// ---- VISUs/Carrousel.TcVIS
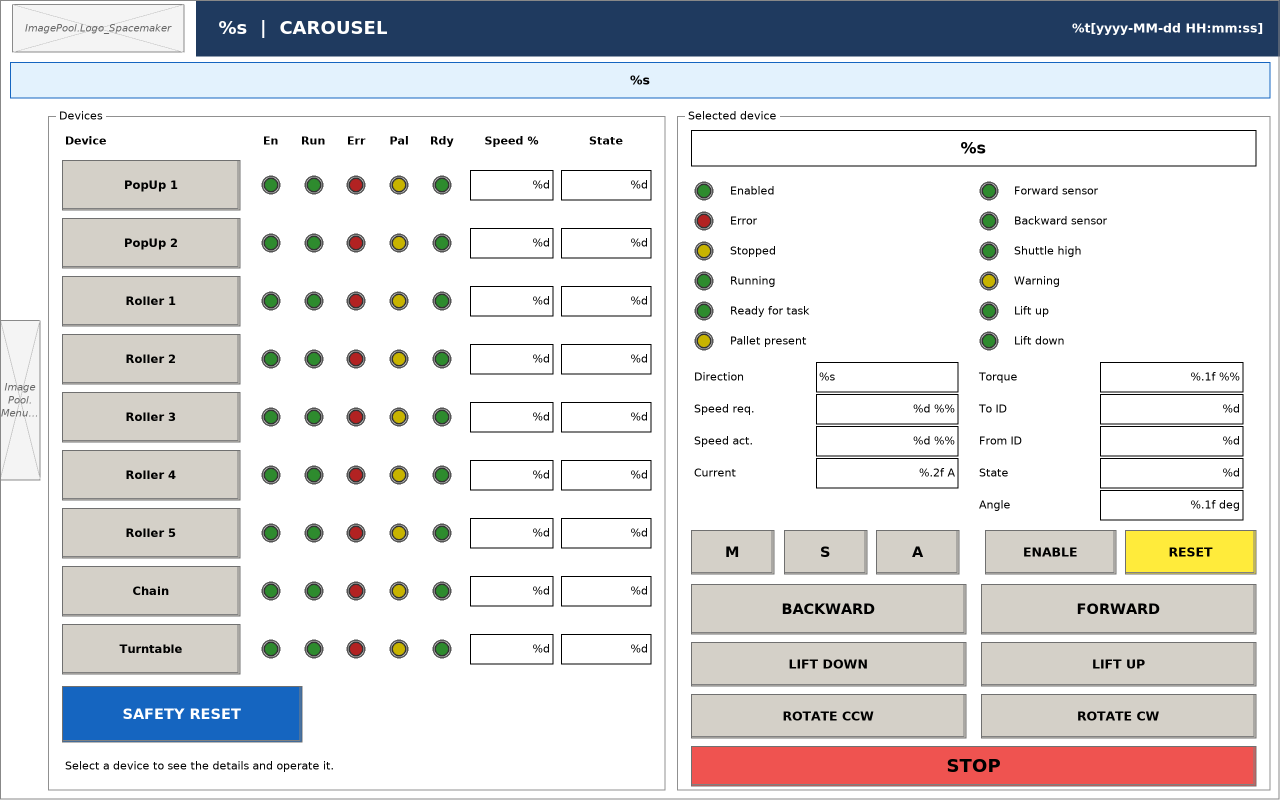
VISUALIZATION Carrousel  // 1280x800
    Rectangle (0,0 196x56)
        OnMouseClick: change screen: Main
    Image (12,4 172x48), image: ImagePool.Logo_Spacemaker
        OnMouseClick: change screen: Main
    Rectangle (196,0 1084x56), "%s | CAROUSEL", text variable: GVL_HMI_System.stStatus.sSystemName
    Rectangle (930,8 336x40), "%t[yyyy-MM-dd HH:mm:ss]", text variable: GVL_HMI_System.stStatus.dtNow
    Rectangle (10,62 1260x36), "%s", text variable: GVL_HMI_System.stStatus.sMessage, colour toggle: GVL_HMI_System.stStatus.bMessageAlarm
    GroupBox (48,108 617x682), "Devices"
    Rectangle (62,128 178x26), "Device"
    Rectangle (250,128 42x26), "En"
    Rectangle (292,128 43x26), "Run"
    Rectangle (335,128 43x26), "Err"
    Rectangle (378,128 43x26), "Pal"
    Rectangle (421,128 42x26), "Rdy"
    Rectangle (470,128 83x26), "Speed %"
    Rectangle (561,128 90x26), "State"
    Button (62,160 178x50), "PopUp 1", colour toggle: GVL_HMI_Carousel.astDevice[1].bSelected
        OnMouseClick: execute { GVL_HMI_Carousel.uiSelected := 1; }
    Lamp1 (260,174 22x22), variable: GVL_HMI_Carousel.astDevice[1].bEnabled, style: Lamp-Lamp1-Green
    Lamp1 (303,174 22x22), variable: GVL_HMI_Carousel.astDevice[1].bRunning, style: Lamp-Lamp1-Green
    Lamp1 (345,174 22x22), variable: GVL_HMI_Carousel.astDevice[1].bError, style: Lamp-Lamp1-Red
    Lamp1 (388,174 22x22), variable: GVL_HMI_Carousel.astDevice[1].bOccupied, style: Lamp-Lamp1-Yellow
    Lamp1 (431,174 22x22), variable: GVL_HMI_Carousel.astDevice[1].bReadyForTask, style: Lamp-Lamp1-Green
    Rectangle (470,170 83x30), "%d", text variable: GVL_HMI_Carousel.astDevice[1].iSpeedActual_pct
    Rectangle (561,170 90x30), "%d", text variable: GVL_HMI_Carousel.astDevice[1].uiStateMachine
    Button (62,218 178x50), "PopUp 2", colour toggle: GVL_HMI_Carousel.astDevice[2].bSelected
        OnMouseClick: execute { GVL_HMI_Carousel.uiSelected := 2; }
    Lamp1 (260,232 22x22), variable: GVL_HMI_Carousel.astDevice[2].bEnabled, style: Lamp-Lamp1-Green
    Lamp1 (303,232 22x22), variable: GVL_HMI_Carousel.astDevice[2].bRunning, style: Lamp-Lamp1-Green
    Lamp1 (345,232 22x22), variable: GVL_HMI_Carousel.astDevice[2].bError, style: Lamp-Lamp1-Red
    Lamp1 (388,232 22x22), variable: GVL_HMI_Carousel.astDevice[2].bOccupied, style: Lamp-Lamp1-Yellow
    Lamp1 (431,232 22x22), variable: GVL_HMI_Carousel.astDevice[2].bReadyForTask, style: Lamp-Lamp1-Green
    Rectangle (470,228 83x30), "%d", text variable: GVL_HMI_Carousel.astDevice[2].iSpeedActual_pct
    Rectangle (561,228 90x30), "%d", text variable: GVL_HMI_Carousel.astDevice[2].uiStateMachine
    Button (62,276 178x50), "Roller 1", colour toggle: GVL_HMI_Carousel.astDevice[3].bSelected
        OnMouseClick: execute { GVL_HMI_Carousel.uiSelected := 3; }
    Lamp1 (260,290 22x22), variable: GVL_HMI_Carousel.astDevice[3].bEnabled, style: Lamp-Lamp1-Green
    Lamp1 (303,290 22x22), variable: GVL_HMI_Carousel.astDevice[3].bRunning, style: Lamp-Lamp1-Green
    Lamp1 (345,290 22x22), variable: GVL_HMI_Carousel.astDevice[3].bError, style: Lamp-Lamp1-Red
    Lamp1 (388,290 22x22), variable: GVL_HMI_Carousel.astDevice[3].bOccupied, style: Lamp-Lamp1-Yellow
    Lamp1 (431,290 22x22), variable: GVL_HMI_Carousel.astDevice[3].bReadyForTask, style: Lamp-Lamp1-Green
    Rectangle (470,286 83x30), "%d", text variable: GVL_HMI_Carousel.astDevice[3].iSpeedActual_pct
    Rectangle (561,286 90x30), "%d", text variable: GVL_HMI_Carousel.astDevice[3].uiStateMachine
    Button (62,334 178x50), "Roller 2", colour toggle: GVL_HMI_Carousel.astDevice[4].bSelected
        OnMouseClick: execute { GVL_HMI_Carousel.uiSelected := 4; }
    Lamp1 (260,348 22x22), variable: GVL_HMI_Carousel.astDevice[4].bEnabled, style: Lamp-Lamp1-Green
    Lamp1 (303,348 22x22), variable: GVL_HMI_Carousel.astDevice[4].bRunning, style: Lamp-Lamp1-Green
    Lamp1 (345,348 22x22), variable: GVL_HMI_Carousel.astDevice[4].bError, style: Lamp-Lamp1-Red
    Lamp1 (388,348 22x22), variable: GVL_HMI_Carousel.astDevice[4].bOccupied, style: Lamp-Lamp1-Yellow
    Lamp1 (431,348 22x22), variable: GVL_HMI_Carousel.astDevice[4].bReadyForTask, style: Lamp-Lamp1-Green
    Rectangle (470,344 83x30), "%d", text variable: GVL_HMI_Carousel.astDevice[4].iSpeedActual_pct
    Rectangle (561,344 90x30), "%d", text variable: GVL_HMI_Carousel.astDevice[4].uiStateMachine
    Button (62,392 178x50), "Roller 3", colour toggle: GVL_HMI_Carousel.astDevice[5].bSelected
        OnMouseClick: execute { GVL_HMI_Carousel.uiSelected := 5; }
    Lamp1 (260,406 22x22), variable: GVL_HMI_Carousel.astDevice[5].bEnabled, style: Lamp-Lamp1-Green
    Lamp1 (303,406 22x22), variable: GVL_HMI_Carousel.astDevice[5].bRunning, style: Lamp-Lamp1-Green
    Lamp1 (345,406 22x22), variable: GVL_HMI_Carousel.astDevice[5].bError, style: Lamp-Lamp1-Red
    Lamp1 (388,406 22x22), variable: GVL_HMI_Carousel.astDevice[5].bOccupied, style: Lamp-Lamp1-Yellow
    Lamp1 (431,406 22x22), variable: GVL_HMI_Carousel.astDevice[5].bReadyForTask, style: Lamp-Lamp1-Green
    Rectangle (470,402 83x30), "%d", text variable: GVL_HMI_Carousel.astDevice[5].iSpeedActual_pct
    Rectangle (561,402 90x30), "%d", text variable: GVL_HMI_Carousel.astDevice[5].uiStateMachine
    Button (62,450 178x50), "Roller 4", colour toggle: GVL_HMI_Carousel.astDevice[6].bSelected
        OnMouseClick: execute { GVL_HMI_Carousel.uiSelected := 6; }
    Lamp1 (260,464 22x22), variable: GVL_HMI_Carousel.astDevice[6].bEnabled, style: Lamp-Lamp1-Green
    Lamp1 (303,464 22x22), variable: GVL_HMI_Carousel.astDevice[6].bRunning, style: Lamp-Lamp1-Green
    Lamp1 (345,464 22x22), variable: GVL_HMI_Carousel.astDevice[6].bError, style: Lamp-Lamp1-Red
    Lamp1 (388,464 22x22), variable: GVL_HMI_Carousel.astDevice[6].bOccupied, style: Lamp-Lamp1-Yellow
    Lamp1 (431,464 22x22), variable: GVL_HMI_Carousel.astDevice[6].bReadyForTask, style: Lamp-Lamp1-Green
    Rectangle (470,460 83x30), "%d", text variable: GVL_HMI_Carousel.astDevice[6].iSpeedActual_pct
    Rectangle (561,460 90x30), "%d", text variable: GVL_HMI_Carousel.astDevice[6].uiStateMachine
    Button (62,508 178x50), "Roller 5", colour toggle: GVL_HMI_Carousel.astDevice[7].bSelected
        OnMouseClick: execute { GVL_HMI_Carousel.uiSelected := 7; }
    Lamp1 (260,522 22x22), variable: GVL_HMI_Carousel.astDevice[7].bEnabled, style: Lamp-Lamp1-Green
    Lamp1 (303,522 22x22), variable: GVL_HMI_Carousel.astDevice[7].bRunning, style: Lamp-Lamp1-Green
    Lamp1 (345,522 22x22), variable: GVL_HMI_Carousel.astDevice[7].bError, style: Lamp-Lamp1-Red
    Lamp1 (388,522 22x22), variable: GVL_HMI_Carousel.astDevice[7].bOccupied, style: Lamp-Lamp1-Yellow
    Lamp1 (431,522 22x22), variable: GVL_HMI_Carousel.astDevice[7].bReadyForTask, style: Lamp-Lamp1-Green
    Rectangle (470,518 83x30), "%d", text variable: GVL_HMI_Carousel.astDevice[7].iSpeedActual_pct
    Rectangle (561,518 90x30), "%d", text variable: GVL_HMI_Carousel.astDevice[7].uiStateMachine
    Button (62,566 178x50), "Chain", colour toggle: GVL_HMI_Carousel.astDevice[8].bSelected
        OnMouseClick: execute { GVL_HMI_Carousel.uiSelected := 8; }
    Lamp1 (260,580 22x22), variable: GVL_HMI_Carousel.astDevice[8].bEnabled, style: Lamp-Lamp1-Green
    Lamp1 (303,580 22x22), variable: GVL_HMI_Carousel.astDevice[8].bRunning, style: Lamp-Lamp1-Green
    Lamp1 (345,580 22x22), variable: GVL_HMI_Carousel.astDevice[8].bError, style: Lamp-Lamp1-Red
    Lamp1 (388,580 22x22), variable: GVL_HMI_Carousel.astDevice[8].bOccupied, style: Lamp-Lamp1-Yellow
    Lamp1 (431,580 22x22), variable: GVL_HMI_Carousel.astDevice[8].bReadyForTask, style: Lamp-Lamp1-Green
    Rectangle (470,576 83x30), "%d", text variable: GVL_HMI_Carousel.astDevice[8].iSpeedActual_pct
    Rectangle (561,576 90x30), "%d", text variable: GVL_HMI_Carousel.astDevice[8].uiStateMachine
    Button (62,624 178x50), "Turntable", colour toggle: GVL_HMI_Carousel.astDevice[9].bSelected
        OnMouseClick: execute { GVL_HMI_Carousel.uiSelected := 9; }
    Lamp1 (260,638 22x22), variable: GVL_HMI_Carousel.astDevice[9].bEnabled, style: Lamp-Lamp1-Green
    Lamp1 (303,638 22x22), variable: GVL_HMI_Carousel.astDevice[9].bRunning, style: Lamp-Lamp1-Green
    Lamp1 (345,638 22x22), variable: GVL_HMI_Carousel.astDevice[9].bError, style: Lamp-Lamp1-Red
    Lamp1 (388,638 22x22), variable: GVL_HMI_Carousel.astDevice[9].bOccupied, style: Lamp-Lamp1-Yellow
    Lamp1 (431,638 22x22), variable: GVL_HMI_Carousel.astDevice[9].bReadyForTask, style: Lamp-Lamp1-Green
    Rectangle (470,634 83x30), "%d", text variable: GVL_HMI_Carousel.astDevice[9].iSpeedActual_pct
    Rectangle (561,634 90x30), "%d", text variable: GVL_HMI_Carousel.astDevice[9].uiStateMachine
    Rectangle (62,752 593x28), "Select a device to see the details and operate it."
    GroupBox (677,108 593x682), "Selected device"
    Rectangle (691,130 565x36), "%s", text variable: GVL_HMI_Carousel.stSelected.sName
    Lamp1 (693,180 22x22), variable: GVL_HMI_Carousel.stSelected.bEnabled, style: Lamp-Lamp1-Green
    Rectangle (727,176 201x30), "Enabled"
    Lamp1 (693,210 22x22), variable: GVL_HMI_Carousel.stSelected.bError, style: Lamp-Lamp1-Red
    Rectangle (727,206 201x30), "Error"
    Lamp1 (693,240 22x22), variable: GVL_HMI_Carousel.stSelected.bStopped, style: Lamp-Lamp1-Yellow
    Rectangle (727,236 201x30), "Stopped"
    Lamp1 (693,270 22x22), variable: GVL_HMI_Carousel.stSelected.bRunning, style: Lamp-Lamp1-Green
    Rectangle (727,266 201x30), "Running"
    Lamp1 (693,300 22x22), variable: GVL_HMI_Carousel.stSelected.bReadyForTask, style: Lamp-Lamp1-Green
    Rectangle (727,296 201x30), "Ready for task"
    Lamp1 (693,330 22x22), variable: GVL_HMI_Carousel.stSelected.bOccupied, style: Lamp-Lamp1-Yellow
    Rectangle (727,326 201x30), "Pallet present"
    Lamp1 (978,180 22x22), variable: GVL_HMI_Carousel.stSelected.bForwardSensor, style: Lamp-Lamp1-Green
    Rectangle (1011,176 202x30), "Forward sensor"
    Lamp1 (978,210 22x22), variable: GVL_HMI_Carousel.stSelected.bBackwardSensor, style: Lamp-Lamp1-Green
    Rectangle (1011,206 202x30), "Backward sensor"
    Lamp1 (978,240 22x22), variable: GVL_HMI_Carousel.stSelected.bShuttleHigh, style: Lamp-Lamp1-Green
    Rectangle (1011,236 202x30), "Shuttle high"
    Lamp1 (978,270 22x22), variable: GVL_HMI_Carousel.stSelected.bWarning, style: Lamp-Lamp1-Yellow
    Rectangle (1011,266 202x30), "Warning"
    Lamp1 (978,300 22x22), variable: GVL_HMI_Carousel.stSelected.bLiftUp, style: Lamp-Lamp1-Green
    Rectangle (1011,296 202x30), "Lift up"
    Lamp1 (978,330 22x22), variable: GVL_HMI_Carousel.stSelected.bLiftDown, style: Lamp-Lamp1-Green
    Rectangle (1011,326 202x30), "Lift down"
    Rectangle (691,362 119x30), "Direction"
    Rectangle (816,362 142x30), "%s", text variable: GVL_HMI_Carousel.stSelected.sMotorDirection
    Rectangle (691,394 119x30), "Speed req."
    Rectangle (816,394 142x30), "%d %%", text variable: GVL_HMI_Carousel.stSelected.iSpeedRequested_pct
    Rectangle (691,426 119x30), "Speed act."
    Rectangle (816,426 142x30), "%d %%", text variable: GVL_HMI_Carousel.stSelected.iSpeedActual_pct
    Rectangle (691,458 119x30), "Current"
    Rectangle (816,458 142x30), "%.2f A", text variable: GVL_HMI_Carousel.stSelected.rCurrent_A
    Rectangle (976,362 118x30), "Torque"
    Rectangle (1100,362 143x30), "%.1f %%", text variable: GVL_HMI_Carousel.stSelected.rTorque_pct
    Rectangle (976,394 118x30), "To ID"
    Rectangle (1100,394 143x30), "%d", text variable: GVL_HMI_Carousel.stSelected.diTransferToId
    Rectangle (976,426 118x30), "From ID"
    Rectangle (1100,426 143x30), "%d", text variable: GVL_HMI_Carousel.stSelected.diTransferFromId
    Rectangle (976,458 118x30), "State"
    Rectangle (1100,458 143x30), "%d", text variable: GVL_HMI_Carousel.stSelected.uiStateMachine
    Rectangle (976,490 118x30), "Angle"
    Rectangle (1100,490 143x30), "%.1f deg", text variable: GVL_HMI_Carousel.stSelected.rAngle_deg
    Button (691,530 83x44), "M", colour toggle: GVL_HMI_Carousel.stSelected.bModeManual
        tap GVL_HMI_Carousel.stCommand.bModeManual p3779583253=TRUE
    Button (784,530 83x44), "S", colour toggle: GVL_HMI_Carousel.stSelected.bModeSemi
        tap GVL_HMI_Carousel.stCommand.bModeSemi p3779583253=TRUE
    Button (876,530 83x44), "A", colour toggle: GVL_HMI_Carousel.stSelected.bModeAuto
        tap GVL_HMI_Carousel.stCommand.bModeAuto p3779583253=TRUE
    Button (985,530 131x44), "ENABLE", colour toggle: GVL_HMI_Carousel.stSelected.bEnabled
        tap GVL_HMI_Carousel.stCommand.bEnable p3779583253=TRUE
    Button (1125,530 131x44), "RESET"
        tap GVL_HMI_Carousel.stCommand.bReset p3779583253=TRUE
    Button (691,584 275x50), "BACKWARD", input disabled if: NOT GVL_HMI_Carousel.stSelected.bModeManual
        tap GVL_HMI_Carousel.stCommand.bJogBackward p3779583253=TRUE
    Button (981,584 275x50), "FORWARD", input disabled if: NOT GVL_HMI_Carousel.stSelected.bModeManual
        tap GVL_HMI_Carousel.stCommand.bJogForward p3779583253=TRUE
    Button (691,642 275x44), "LIFT DOWN", input disabled if: NOT GVL_HMI_Carousel.stSelected.bHasLift
        tap GVL_HMI_Carousel.stCommand.bLiftDown p3779583253=TRUE
    Button (981,642 275x44), "LIFT UP", input disabled if: NOT GVL_HMI_Carousel.stSelected.bHasLift
        tap GVL_HMI_Carousel.stCommand.bLiftUp p3779583253=TRUE
    Button (691,694 275x44), "ROTATE CCW", input disabled if: NOT GVL_HMI_Carousel.stSelected.bHasRotation
        tap GVL_HMI_Carousel.stCommand.bRotateCcw p3779583253=TRUE
    Button (981,694 275x44), "ROTATE CW", input disabled if: NOT GVL_HMI_Carousel.stSelected.bHasRotation
        tap GVL_HMI_Carousel.stCommand.bRotateCw p3779583253=TRUE
    Button (691,746 565x40), "STOP"
        tap GVL_HMI_Carousel.stCommand.bStop p3779583253=TRUE
    Rectangle (0,320 40x160)
        OnMouseClick: OpenDialog Dialog=Dialog, OpenModal=True, PositionX=0, PositionY=0
        OnMouseEnter: OpenDialog Dialog=Dialog, OpenModal=True, PositionX=0, PositionY=0
    Image (0,320 40x160), image: ImagePool.Menu_Tab
        OnMouseClick: OpenDialog Dialog=Dialog, OpenModal=True, PositionX=0, PositionY=0
        OnMouseEnter: OpenDialog Dialog=Dialog, OpenModal=True, PositionX=0, PositionY=0
    Button (62,686 240x56), "SAFETY RESET", colour toggle: GVL_HMI_System.stStatus.bSafetyResetActive
        tap GVL_HMI_System.stCommand.bSafetyReset p3779583253=TRUE
END_VISUALIZATION

// ---- VISUs/CNV.TcVIS
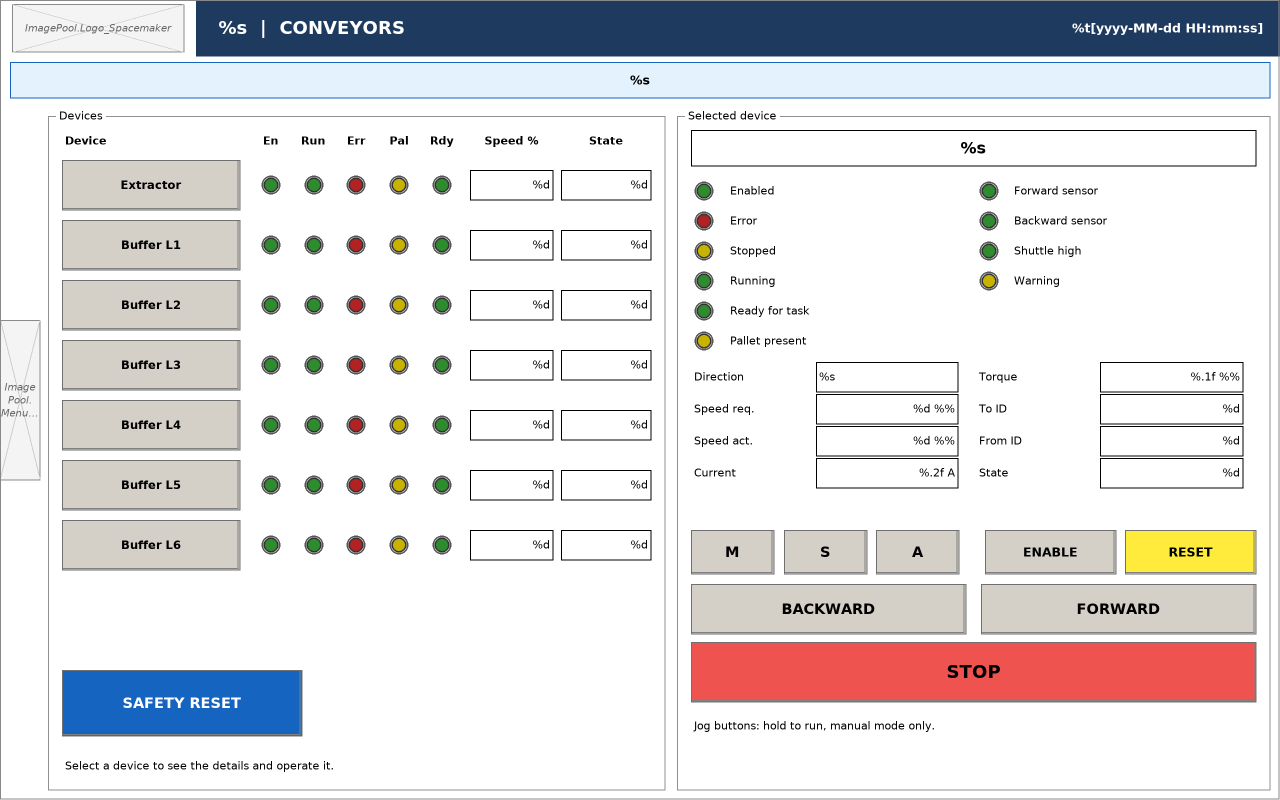
VISUALIZATION CNV  // 1280x800
    Rectangle (0,0 196x56)
        OnMouseClick: change screen: Main
    Image (12,4 172x48), image: ImagePool.Logo_Spacemaker
        OnMouseClick: change screen: Main
    Rectangle (196,0 1084x56), "%s | CONVEYORS", text variable: GVL_HMI_System.stStatus.sSystemName
    Rectangle (930,8 336x40), "%t[yyyy-MM-dd HH:mm:ss]", text variable: GVL_HMI_System.stStatus.dtNow
    Rectangle (10,62 1260x36), "%s", text variable: GVL_HMI_System.stStatus.sMessage, colour toggle: GVL_HMI_System.stStatus.bMessageAlarm
    GroupBox (48,108 617x682), "Devices"
    Rectangle (62,128 178x26), "Device"
    Rectangle (250,128 42x26), "En"
    Rectangle (292,128 43x26), "Run"
    Rectangle (335,128 43x26), "Err"
    Rectangle (378,128 43x26), "Pal"
    Rectangle (421,128 42x26), "Rdy"
    Rectangle (470,128 83x26), "Speed %"
    Rectangle (561,128 90x26), "State"
    Button (62,160 178x50), "Extractor", colour toggle: GVL_HMI_CNV.astConveyor[0].bSelected
        OnMouseClick: execute { GVL_HMI_CNV.uiSelected := 0; }
    Lamp1 (260,174 22x22), variable: GVL_HMI_CNV.astConveyor[0].bEnabled, style: Lamp-Lamp1-Green
    Lamp1 (303,174 22x22), variable: GVL_HMI_CNV.astConveyor[0].bRunning, style: Lamp-Lamp1-Green
    Lamp1 (345,174 22x22), variable: GVL_HMI_CNV.astConveyor[0].bError, style: Lamp-Lamp1-Red
    Lamp1 (388,174 22x22), variable: GVL_HMI_CNV.astConveyor[0].bOccupied, style: Lamp-Lamp1-Yellow
    Lamp1 (431,174 22x22), variable: GVL_HMI_CNV.astConveyor[0].bReadyForTask, style: Lamp-Lamp1-Green
    Rectangle (470,170 83x30), "%d", text variable: GVL_HMI_CNV.astConveyor[0].iSpeedActual_pct
    Rectangle (561,170 90x30), "%d", text variable: GVL_HMI_CNV.astConveyor[0].uiStateMachine
    Button (62,220 178x50), "Buffer L1", colour toggle: GVL_HMI_CNV.astConveyor[1].bSelected
        OnMouseClick: execute { GVL_HMI_CNV.uiSelected := 1; }
    Lamp1 (260,234 22x22), variable: GVL_HMI_CNV.astConveyor[1].bEnabled, style: Lamp-Lamp1-Green
    Lamp1 (303,234 22x22), variable: GVL_HMI_CNV.astConveyor[1].bRunning, style: Lamp-Lamp1-Green
    Lamp1 (345,234 22x22), variable: GVL_HMI_CNV.astConveyor[1].bError, style: Lamp-Lamp1-Red
    Lamp1 (388,234 22x22), variable: GVL_HMI_CNV.astConveyor[1].bOccupied, style: Lamp-Lamp1-Yellow
    Lamp1 (431,234 22x22), variable: GVL_HMI_CNV.astConveyor[1].bReadyForTask, style: Lamp-Lamp1-Green
    Rectangle (470,230 83x30), "%d", text variable: GVL_HMI_CNV.astConveyor[1].iSpeedActual_pct
    Rectangle (561,230 90x30), "%d", text variable: GVL_HMI_CNV.astConveyor[1].uiStateMachine
    Button (62,280 178x50), "Buffer L2", colour toggle: GVL_HMI_CNV.astConveyor[2].bSelected
        OnMouseClick: execute { GVL_HMI_CNV.uiSelected := 2; }
    Lamp1 (260,294 22x22), variable: GVL_HMI_CNV.astConveyor[2].bEnabled, style: Lamp-Lamp1-Green
    Lamp1 (303,294 22x22), variable: GVL_HMI_CNV.astConveyor[2].bRunning, style: Lamp-Lamp1-Green
    Lamp1 (345,294 22x22), variable: GVL_HMI_CNV.astConveyor[2].bError, style: Lamp-Lamp1-Red
    Lamp1 (388,294 22x22), variable: GVL_HMI_CNV.astConveyor[2].bOccupied, style: Lamp-Lamp1-Yellow
    Lamp1 (431,294 22x22), variable: GVL_HMI_CNV.astConveyor[2].bReadyForTask, style: Lamp-Lamp1-Green
    Rectangle (470,290 83x30), "%d", text variable: GVL_HMI_CNV.astConveyor[2].iSpeedActual_pct
    Rectangle (561,290 90x30), "%d", text variable: GVL_HMI_CNV.astConveyor[2].uiStateMachine
    Button (62,340 178x50), "Buffer L3", colour toggle: GVL_HMI_CNV.astConveyor[3].bSelected
        OnMouseClick: execute { GVL_HMI_CNV.uiSelected := 3; }
    Lamp1 (260,354 22x22), variable: GVL_HMI_CNV.astConveyor[3].bEnabled, style: Lamp-Lamp1-Green
    Lamp1 (303,354 22x22), variable: GVL_HMI_CNV.astConveyor[3].bRunning, style: Lamp-Lamp1-Green
    Lamp1 (345,354 22x22), variable: GVL_HMI_CNV.astConveyor[3].bError, style: Lamp-Lamp1-Red
    Lamp1 (388,354 22x22), variable: GVL_HMI_CNV.astConveyor[3].bOccupied, style: Lamp-Lamp1-Yellow
    Lamp1 (431,354 22x22), variable: GVL_HMI_CNV.astConveyor[3].bReadyForTask, style: Lamp-Lamp1-Green
    Rectangle (470,350 83x30), "%d", text variable: GVL_HMI_CNV.astConveyor[3].iSpeedActual_pct
    Rectangle (561,350 90x30), "%d", text variable: GVL_HMI_CNV.astConveyor[3].uiStateMachine
    Button (62,400 178x50), "Buffer L4", colour toggle: GVL_HMI_CNV.astConveyor[4].bSelected
        OnMouseClick: execute { GVL_HMI_CNV.uiSelected := 4; }
    Lamp1 (260,414 22x22), variable: GVL_HMI_CNV.astConveyor[4].bEnabled, style: Lamp-Lamp1-Green
    Lamp1 (303,414 22x22), variable: GVL_HMI_CNV.astConveyor[4].bRunning, style: Lamp-Lamp1-Green
    Lamp1 (345,414 22x22), variable: GVL_HMI_CNV.astConveyor[4].bError, style: Lamp-Lamp1-Red
    Lamp1 (388,414 22x22), variable: GVL_HMI_CNV.astConveyor[4].bOccupied, style: Lamp-Lamp1-Yellow
    Lamp1 (431,414 22x22), variable: GVL_HMI_CNV.astConveyor[4].bReadyForTask, style: Lamp-Lamp1-Green
    Rectangle (470,410 83x30), "%d", text variable: GVL_HMI_CNV.astConveyor[4].iSpeedActual_pct
    Rectangle (561,410 90x30), "%d", text variable: GVL_HMI_CNV.astConveyor[4].uiStateMachine
    Button (62,460 178x50), "Buffer L5", colour toggle: GVL_HMI_CNV.astConveyor[5].bSelected
        OnMouseClick: execute { GVL_HMI_CNV.uiSelected := 5; }
    Lamp1 (260,474 22x22), variable: GVL_HMI_CNV.astConveyor[5].bEnabled, style: Lamp-Lamp1-Green
    Lamp1 (303,474 22x22), variable: GVL_HMI_CNV.astConveyor[5].bRunning, style: Lamp-Lamp1-Green
    Lamp1 (345,474 22x22), variable: GVL_HMI_CNV.astConveyor[5].bError, style: Lamp-Lamp1-Red
    Lamp1 (388,474 22x22), variable: GVL_HMI_CNV.astConveyor[5].bOccupied, style: Lamp-Lamp1-Yellow
    Lamp1 (431,474 22x22), variable: GVL_HMI_CNV.astConveyor[5].bReadyForTask, style: Lamp-Lamp1-Green
    Rectangle (470,470 83x30), "%d", text variable: GVL_HMI_CNV.astConveyor[5].iSpeedActual_pct
    Rectangle (561,470 90x30), "%d", text variable: GVL_HMI_CNV.astConveyor[5].uiStateMachine
    Button (62,520 178x50), "Buffer L6", colour toggle: GVL_HMI_CNV.astConveyor[6].bSelected
        OnMouseClick: execute { GVL_HMI_CNV.uiSelected := 6; }
    Lamp1 (260,534 22x22), variable: GVL_HMI_CNV.astConveyor[6].bEnabled, style: Lamp-Lamp1-Green
    Lamp1 (303,534 22x22), variable: GVL_HMI_CNV.astConveyor[6].bRunning, style: Lamp-Lamp1-Green
    Lamp1 (345,534 22x22), variable: GVL_HMI_CNV.astConveyor[6].bError, style: Lamp-Lamp1-Red
    Lamp1 (388,534 22x22), variable: GVL_HMI_CNV.astConveyor[6].bOccupied, style: Lamp-Lamp1-Yellow
    Lamp1 (431,534 22x22), variable: GVL_HMI_CNV.astConveyor[6].bReadyForTask, style: Lamp-Lamp1-Green
    Rectangle (470,530 83x30), "%d", text variable: GVL_HMI_CNV.astConveyor[6].iSpeedActual_pct
    Rectangle (561,530 90x30), "%d", text variable: GVL_HMI_CNV.astConveyor[6].uiStateMachine
    Rectangle (62,752 593x28), "Select a device to see the details and operate it."
    GroupBox (677,108 593x682), "Selected device"
    Rectangle (691,130 565x36), "%s", text variable: GVL_HMI_CNV.stSelected.sName
    Lamp1 (693,180 22x22), variable: GVL_HMI_CNV.stSelected.bEnabled, style: Lamp-Lamp1-Green
    Rectangle (727,176 201x30), "Enabled"
    Lamp1 (693,210 22x22), variable: GVL_HMI_CNV.stSelected.bError, style: Lamp-Lamp1-Red
    Rectangle (727,206 201x30), "Error"
    Lamp1 (693,240 22x22), variable: GVL_HMI_CNV.stSelected.bStopped, style: Lamp-Lamp1-Yellow
    Rectangle (727,236 201x30), "Stopped"
    Lamp1 (693,270 22x22), variable: GVL_HMI_CNV.stSelected.bRunning, style: Lamp-Lamp1-Green
    Rectangle (727,266 201x30), "Running"
    Lamp1 (693,300 22x22), variable: GVL_HMI_CNV.stSelected.bReadyForTask, style: Lamp-Lamp1-Green
    Rectangle (727,296 201x30), "Ready for task"
    Lamp1 (693,330 22x22), variable: GVL_HMI_CNV.stSelected.bOccupied, style: Lamp-Lamp1-Yellow
    Rectangle (727,326 201x30), "Pallet present"
    Lamp1 (978,180 22x22), variable: GVL_HMI_CNV.stSelected.bForwardSensor, style: Lamp-Lamp1-Green
    Rectangle (1011,176 202x30), "Forward sensor"
    Lamp1 (978,210 22x22), variable: GVL_HMI_CNV.stSelected.bBackwardSensor, style: Lamp-Lamp1-Green
    Rectangle (1011,206 202x30), "Backward sensor"
    Lamp1 (978,240 22x22), variable: GVL_HMI_CNV.stSelected.bShuttleHigh, style: Lamp-Lamp1-Green
    Rectangle (1011,236 202x30), "Shuttle high"
    Lamp1 (978,270 22x22), variable: GVL_HMI_CNV.stSelected.bWarning, style: Lamp-Lamp1-Yellow
    Rectangle (1011,266 202x30), "Warning"
    Rectangle (691,362 119x30), "Direction"
    Rectangle (816,362 142x30), "%s", text variable: GVL_HMI_CNV.stSelected.sMotorDirection
    Rectangle (691,394 119x30), "Speed req."
    Rectangle (816,394 142x30), "%d %%", text variable: GVL_HMI_CNV.stSelected.iSpeedRequested_pct
    Rectangle (691,426 119x30), "Speed act."
    Rectangle (816,426 142x30), "%d %%", text variable: GVL_HMI_CNV.stSelected.iSpeedActual_pct
    Rectangle (691,458 119x30), "Current"
    Rectangle (816,458 142x30), "%.2f A", text variable: GVL_HMI_CNV.stSelected.rCurrent_A
    Rectangle (976,362 118x30), "Torque"
    Rectangle (1100,362 143x30), "%.1f %%", text variable: GVL_HMI_CNV.stSelected.rTorque_pct
    Rectangle (976,394 118x30), "To ID"
    Rectangle (1100,394 143x30), "%d", text variable: GVL_HMI_CNV.stSelected.diTransferToId
    Rectangle (976,426 118x30), "From ID"
    Rectangle (1100,426 143x30), "%d", text variable: GVL_HMI_CNV.stSelected.diTransferFromId
    Rectangle (976,458 118x30), "State"
    Rectangle (1100,458 143x30), "%d", text variable: GVL_HMI_CNV.stSelected.uiStateMachine
    Button (691,530 83x44), "M", colour toggle: GVL_HMI_CNV.stSelected.bModeManual
        tap GVL_HMI_CNV.stCommand.bModeManual p3779583253=TRUE
    Button (784,530 83x44), "S", colour toggle: GVL_HMI_CNV.stSelected.bModeSemi
        tap GVL_HMI_CNV.stCommand.bModeSemi p3779583253=TRUE
    Button (876,530 83x44), "A", colour toggle: GVL_HMI_CNV.stSelected.bModeAuto
        tap GVL_HMI_CNV.stCommand.bModeAuto p3779583253=TRUE
    Button (985,530 131x44), "ENABLE", colour toggle: GVL_HMI_CNV.stSelected.bEnabled
        tap GVL_HMI_CNV.stCommand.bEnable p3779583253=TRUE
    Button (1125,530 131x44), "RESET"
        tap GVL_HMI_CNV.stCommand.bReset p3779583253=TRUE
    Button (691,584 275x50), "BACKWARD", input disabled if: NOT GVL_HMI_CNV.stSelected.bModeManual
        tap GVL_HMI_CNV.stCommand.bJogBackward p3779583253=TRUE
    Button (981,584 275x50), "FORWARD", input disabled if: NOT GVL_HMI_CNV.stSelected.bModeManual
        tap GVL_HMI_CNV.stCommand.bJogForward p3779583253=TRUE
    Button (691,642 565x60), "STOP"
        tap GVL_HMI_CNV.stCommand.bStop p3779583253=TRUE
    Rectangle (691,712 565x28), "Jog buttons: hold to run, manual mode only."
    Rectangle (0,320 40x160)
        OnMouseClick: OpenDialog Dialog=Dialog, OpenModal=True, PositionX=0, PositionY=0
        OnMouseEnter: OpenDialog Dialog=Dialog, OpenModal=True, PositionX=0, PositionY=0
    Image (0,320 40x160), image: ImagePool.Menu_Tab
        OnMouseClick: OpenDialog Dialog=Dialog, OpenModal=True, PositionX=0, PositionY=0
        OnMouseEnter: OpenDialog Dialog=Dialog, OpenModal=True, PositionX=0, PositionY=0
    Button (62,670 240x66), "SAFETY RESET", colour toggle: GVL_HMI_System.stStatus.bSafetyResetActive
        tap GVL_HMI_System.stCommand.bSafetyReset p3779583253=TRUE
END_VISUALIZATION

// ---- VISUs/CNV_Settings.TcVIS
VISUALIZATION CNV_Settings  // 1024x768
END_VISUALIZATION

// ---- VISUs/Dialog.TcVIS
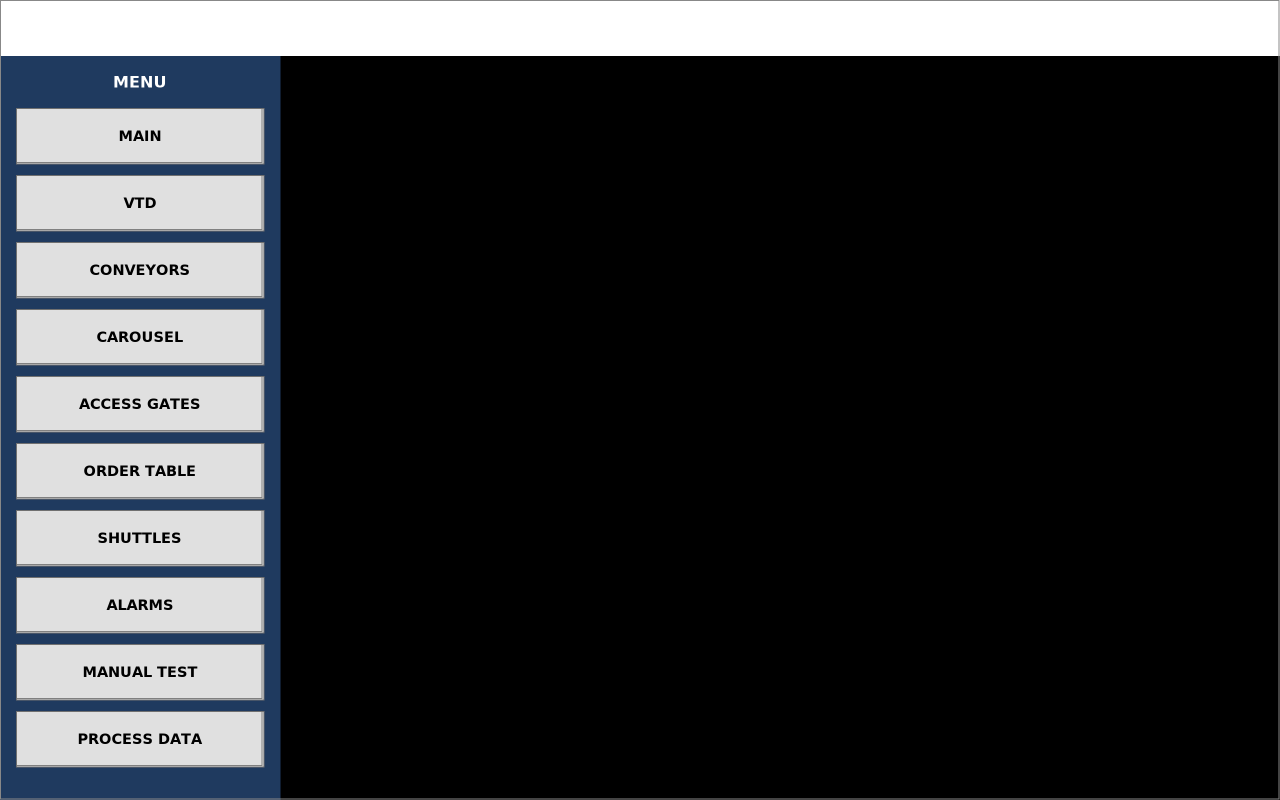
VISUALIZATION Dialog  // 1280x800
    Rectangle (0,0 1280x56)
        OnMouseClick: CloseDialog Dialog=Current Dialog, Result=OK, NumpadKeypadSet=True
    Rectangle (280,56 1000x744)
        OnMouseClick: CloseDialog Dialog=Current Dialog, Result=OK, NumpadKeypadSet=True
    Rectangle (0,56 280x744)
    Rectangle (12,64 256x36), "MENU"
    Button (16,108 248x56), "MAIN"
        OnMouseClick: CloseDialog Dialog=Current Dialog, Result=OK, NumpadKeypadSet=True
        OnMouseDown: change screen: Main
    Button (16,175 248x56), "VTD"
        OnMouseClick: CloseDialog Dialog=Current Dialog, Result=OK, NumpadKeypadSet=True
        OnMouseDown: change screen: VTD
    Button (16,242 248x56), "CONVEYORS"
        OnMouseClick: CloseDialog Dialog=Current Dialog, Result=OK, NumpadKeypadSet=True
        OnMouseDown: change screen: CNV
    Button (16,309 248x56), "CAROUSEL"
        OnMouseClick: CloseDialog Dialog=Current Dialog, Result=OK, NumpadKeypadSet=True
        OnMouseDown: change screen: Carrousel
    Button (16,376 248x56), "ACCESS GATES"
        OnMouseClick: CloseDialog Dialog=Current Dialog, Result=OK, NumpadKeypadSet=True
        OnMouseDown: change screen: Access_Gates
    Button (16,443 248x56), "ORDER TABLE"
        OnMouseClick: CloseDialog Dialog=Current Dialog, Result=OK, NumpadKeypadSet=True
        OnMouseDown: change screen: Order_Table
    Button (16,510 248x56), "SHUTTLES"
        OnMouseClick: CloseDialog Dialog=Current Dialog, Result=OK, NumpadKeypadSet=True
        OnMouseDown: change screen: Shuttles
    Button (16,577 248x56), "ALARMS"
        OnMouseClick: CloseDialog Dialog=Current Dialog, Result=OK, NumpadKeypadSet=True
        OnMouseDown: change screen: Alarms
    Button (16,644 248x56), "MANUAL TEST"
        OnMouseClick: CloseDialog Dialog=Current Dialog, Result=OK, NumpadKeypadSet=True
        OnMouseDown: change screen: VTDManualTest
    Button (16,711 248x56), "PROCESS DATA"
        OnMouseClick: CloseDialog Dialog=Current Dialog, Result=OK, NumpadKeypadSet=True
        OnMouseDown: change screen: Visualization
END_VISUALIZATION

// ---- VISUs/FP_Conveyor.TcVIS
VISUALIZATION FP_Conveyor  // 2x2
END_VISUALIZATION

// ---- VISUs/FP_Drive.TcVIS
VISUALIZATION FP_Drive  // 1024x768
END_VISUALIZATION

// ---- VISUs/FP_Test.TcVIS
VISUALIZATION FP_Test  // 2x2
VAR_IN_OUT
	bTest : BOOL;
END_VAR
END_VISUALIZATION

// ---- VISUs/Header.TcVIS
VISUALIZATION Header  // 1024x768
END_VISUALIZATION

// ---- VISUs/Main.TcVIS
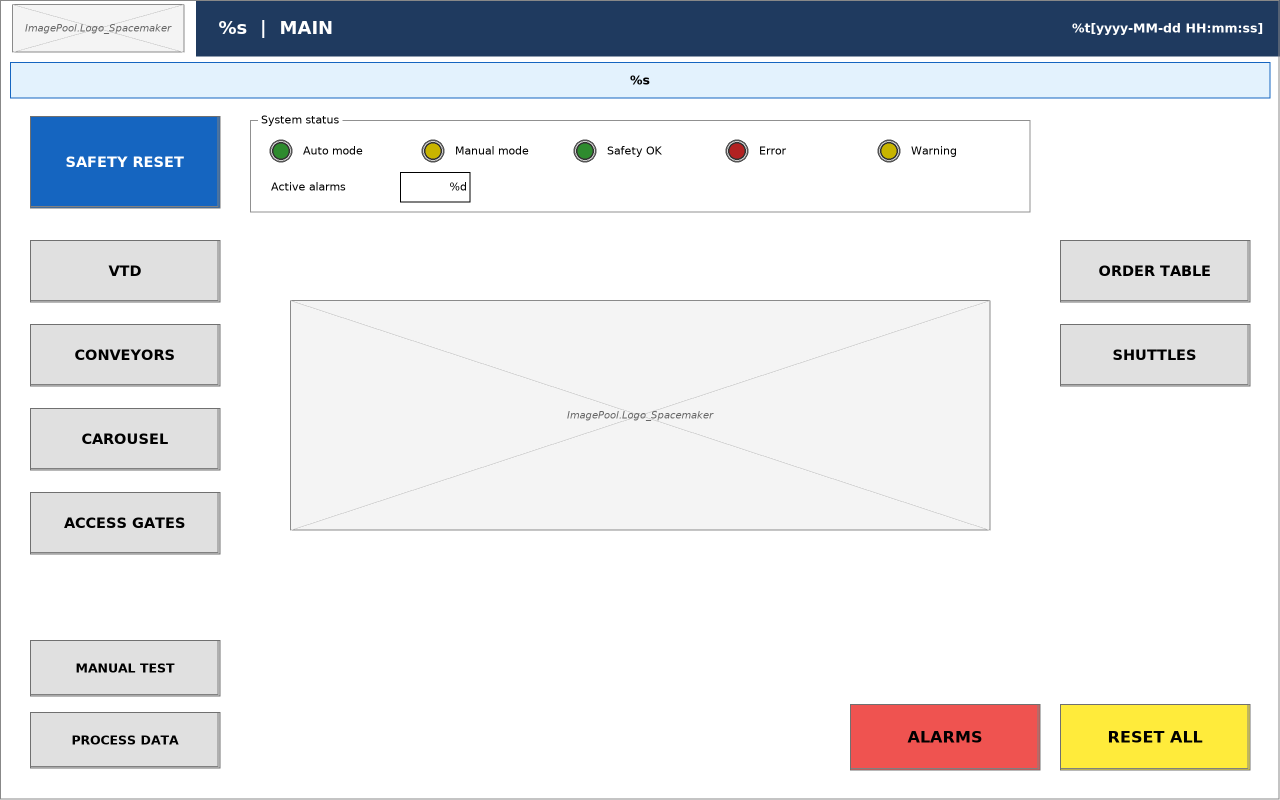
VISUALIZATION Main  // 1280x800
    Rectangle (0,0 196x56)
        OnMouseClick: change screen: Main
    Image (12,4 172x48), image: ImagePool.Logo_Spacemaker
        OnMouseClick: change screen: Main
    Rectangle (196,0 1084x56), "%s | MAIN", text variable: GVL_HMI_System.stStatus.sSystemName
    Rectangle (930,8 336x40), "%t[yyyy-MM-dd HH:mm:ss]", text variable: GVL_HMI_System.stStatus.dtNow
    Rectangle (10,62 1260x36), "%s", text variable: GVL_HMI_System.stStatus.sMessage, colour toggle: GVL_HMI_System.stStatus.bMessageAlarm
    GroupBox (250,112 780x100), "System status"
    Lamp1 (268,138 26x26), variable: GVL_HMI_System.stStatus.bAutoMode, style: Lamp-Lamp1-Green
    Rectangle (300,136 112x30), "Auto mode"
    Lamp1 (420,138 26x26), variable: GVL_HMI_System.stStatus.bManualMode, style: Lamp-Lamp1-Yellow
    Rectangle (452,136 112x30), "Manual mode"
    Lamp1 (572,138 26x26), variable: GVL_HMI_System.stStatus.bSafetyOk, style: Lamp-Lamp1-Green
    Rectangle (604,136 112x30), "Safety OK"
    Lamp1 (724,138 26x26), variable: GVL_HMI_System.stStatus.bError, style: Lamp-Lamp1-Red
    Rectangle (756,136 112x30), "Error"
    Lamp1 (876,138 26x26), variable: GVL_HMI_System.stStatus.bWarning, style: Lamp-Lamp1-Yellow
    Rectangle (908,136 112x30), "Warning"
    Rectangle (268,172 130x30), "Active alarms"
    Rectangle (400,172 70x30), "%d", text variable: GVL_HMI_System.stStatus.uiActiveAlarms
    Image (290,300 700x230), image: ImagePool.Logo_Spacemaker
    Button (30,240 190x62), "VTD", colour toggle: GVL_HMI_System.stVtd.stSummary.bError
        OnMouseClick: change screen: VTD
    Button (30,324 190x62), "CONVEYORS"
        OnMouseClick: change screen: CNV
    Button (30,408 190x62), "CAROUSEL"
        OnMouseClick: change screen: Carrousel
    Button (30,492 190x62), "ACCESS GATES"
        OnMouseClick: change screen: Access_Gates
    Button (30,640 190x56), "MANUAL TEST"
        OnMouseClick: change screen: VTDManualTest
    Button (30,712 190x56), "PROCESS DATA"
        OnMouseClick: change screen: Visualization
    Button (1060,240 190x62), "ORDER TABLE"
        OnMouseClick: change screen: Order_Table
    Button (1060,324 190x62), "SHUTTLES"
        OnMouseClick: change screen: Shuttles
    Button (850,704 190x66), "ALARMS"
        OnMouseClick: change screen: Alarms
    Button (1060,704 190x66), "RESET ALL"
        tap GVL_HMI_System.stCommand.bResetAll p3779583253=TRUE
    Button (30,116 190x92), "SAFETY RESET", colour toggle: GVL_HMI_System.stStatus.bSafetyResetActive
        tap GVL_HMI_System.stCommand.bSafetyReset p3779583253=TRUE
END_VISUALIZATION

// ---- VISUs/NavBar.TcVIS
VISUALIZATION NavBar  // 1024x768
END_VISUALIZATION

// ---- VISUs/Order_Table.TcVIS
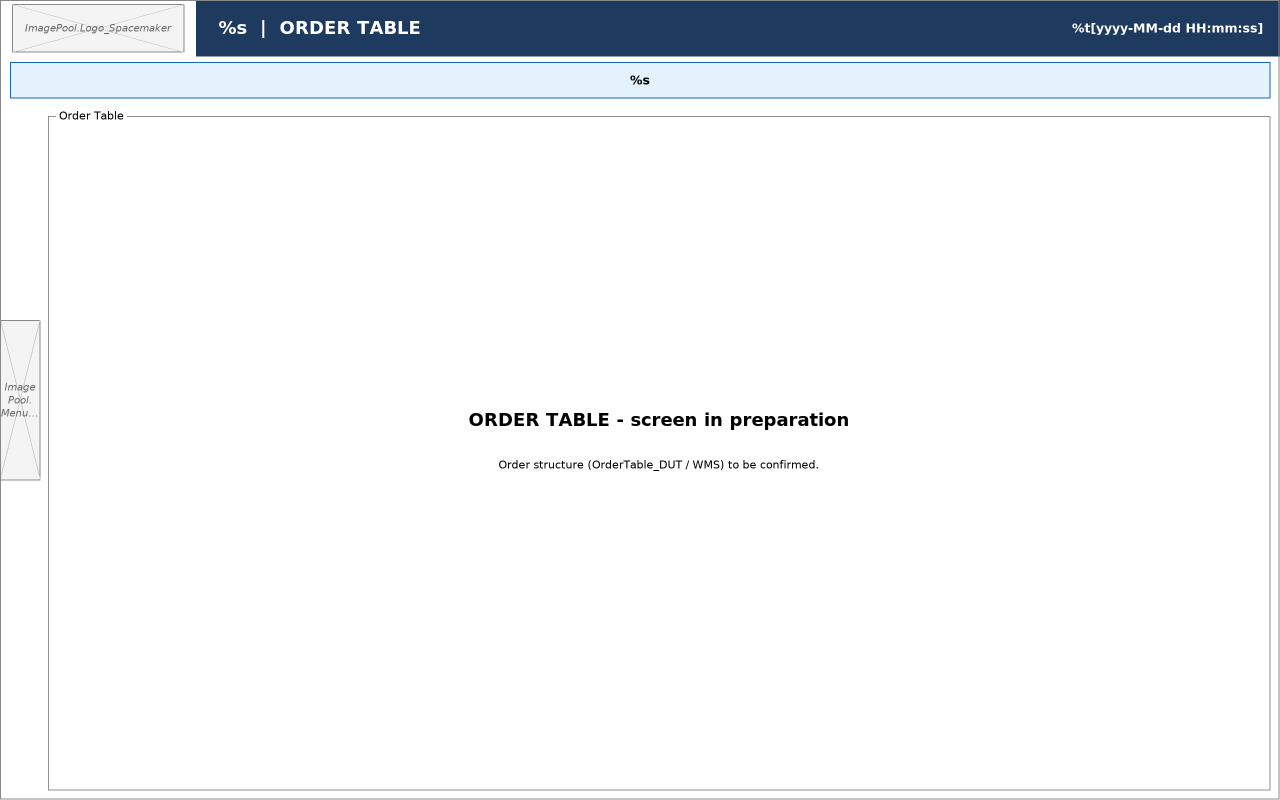
VISUALIZATION Order_Table  // 1280x800
    Rectangle (0,0 196x56)
        OnMouseClick: change screen: Main
    Image (12,4 172x48), image: ImagePool.Logo_Spacemaker
        OnMouseClick: change screen: Main
    Rectangle (196,0 1084x56), "%s | ORDER TABLE", text variable: GVL_HMI_System.stStatus.sSystemName
    Rectangle (930,8 336x40), "%t[yyyy-MM-dd HH:mm:ss]", text variable: GVL_HMI_System.stStatus.dtNow
    Rectangle (10,62 1260x36), "%s", text variable: GVL_HMI_System.stStatus.sMessage, colour toggle: GVL_HMI_System.stStatus.bMessageAlarm
    GroupBox (48,108 1222x682), "Order Table"
    Rectangle (78,400 1162x40), "ORDER TABLE - screen in preparation"
    Rectangle (78,450 1162x30), "Order structure (OrderTable_DUT / WMS) to be confirmed."
    Rectangle (0,320 40x160)
        OnMouseClick: OpenDialog Dialog=Dialog, OpenModal=True, PositionX=0, PositionY=0
        OnMouseEnter: OpenDialog Dialog=Dialog, OpenModal=True, PositionX=0, PositionY=0
    Image (0,320 40x160), image: ImagePool.Menu_Tab
        OnMouseClick: OpenDialog Dialog=Dialog, OpenModal=True, PositionX=0, PositionY=0
        OnMouseEnter: OpenDialog Dialog=Dialog, OpenModal=True, PositionX=0, PositionY=0
END_VISUALIZATION

// ---- VISUs/Shuttles.TcVIS
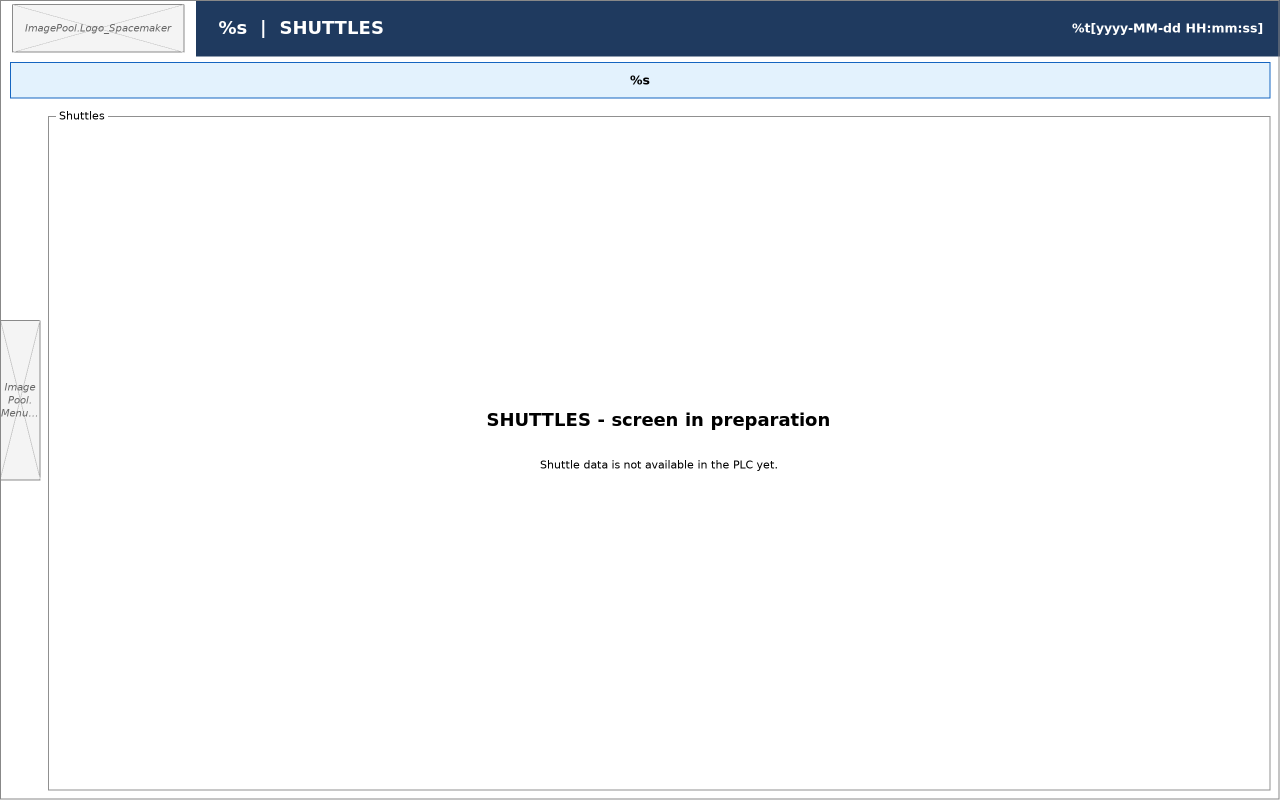
VISUALIZATION Shuttles  // 1280x800
    Rectangle (0,0 196x56)
        OnMouseClick: change screen: Main
    Image (12,4 172x48), image: ImagePool.Logo_Spacemaker
        OnMouseClick: change screen: Main
    Rectangle (196,0 1084x56), "%s | SHUTTLES", text variable: GVL_HMI_System.stStatus.sSystemName
    Rectangle (930,8 336x40), "%t[yyyy-MM-dd HH:mm:ss]", text variable: GVL_HMI_System.stStatus.dtNow
    Rectangle (10,62 1260x36), "%s", text variable: GVL_HMI_System.stStatus.sMessage, colour toggle: GVL_HMI_System.stStatus.bMessageAlarm
    GroupBox (48,108 1222x682), "Shuttles"
    Rectangle (78,400 1162x40), "SHUTTLES - screen in preparation"
    Rectangle (78,450 1162x30), "Shuttle data is not available in the PLC yet."
    Rectangle (0,320 40x160)
        OnMouseClick: OpenDialog Dialog=Dialog, OpenModal=True, PositionX=0, PositionY=0
        OnMouseEnter: OpenDialog Dialog=Dialog, OpenModal=True, PositionX=0, PositionY=0
    Image (0,320 40x160), image: ImagePool.Menu_Tab
        OnMouseClick: OpenDialog Dialog=Dialog, OpenModal=True, PositionX=0, PositionY=0
        OnMouseEnter: OpenDialog Dialog=Dialog, OpenModal=True, PositionX=0, PositionY=0
END_VISUALIZATION

// ---- VISUs/teste.TcVIS
VISUALIZATION teste  // 1024x768
END_VISUALIZATION

// ---- VISUs/Visualization.TcVIS
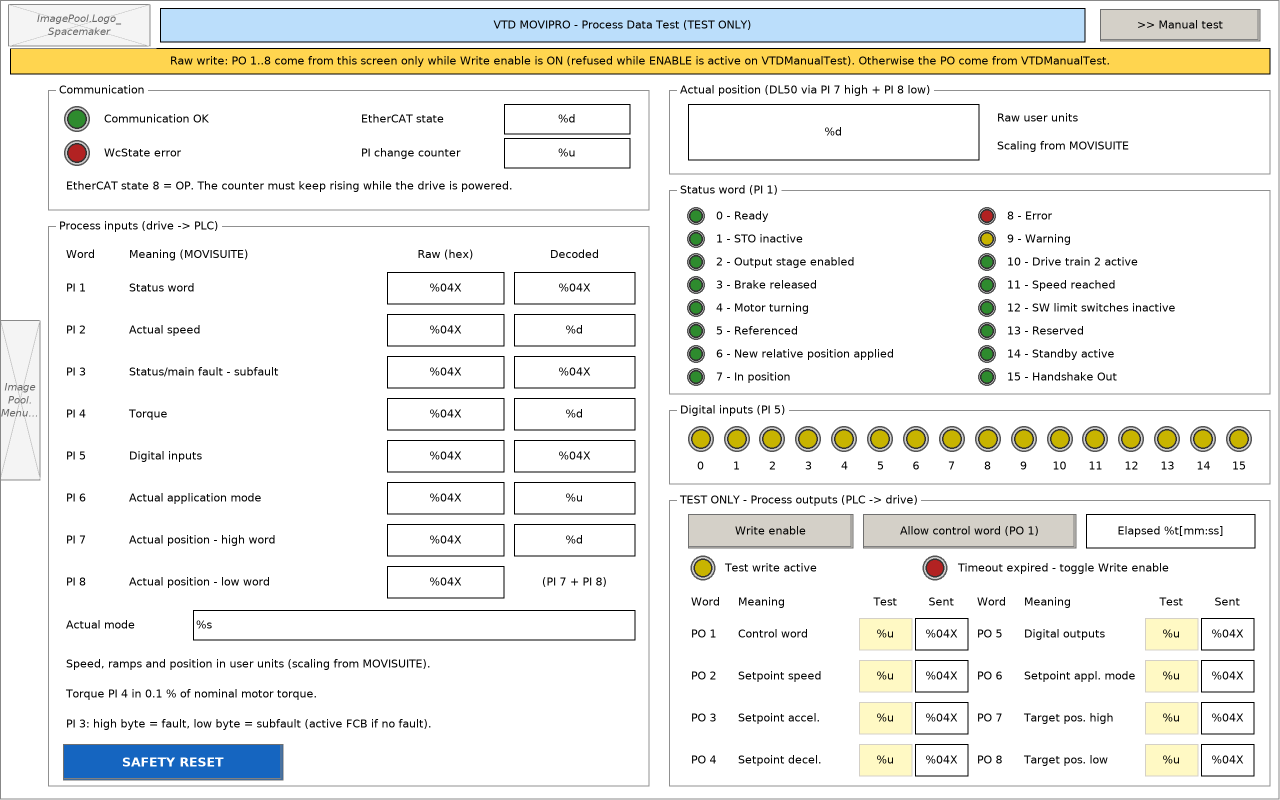
VISUALIZATION Visualization  // 1280x800
    GroupBox (48,82 601x128), "Communication"
    GroupBox (48,218 601x568), "Process inputs (drive -> PLC)"
    GroupBox (669,82 601x92), "Actual position (DL50 via PI 7 high + PI 8 low)"
    GroupBox (669,182 601x212), "Status word (PI 1)"
    GroupBox (669,402 601x82), "Digital inputs (PI 5)"
    GroupBox (669,492 601x294), "TEST ONLY - Process outputs (PLC -> drive)"
    Rectangle (160,8 925x34), "VTD MOVIPRO - Process Data Test (TEST ONLY)"
    Rectangle (10,48 1260x26), "Raw write: PO 1..8 come from this screen only while Write enable is ON (refused while ENABLE is active on VTDManualTest). Otherwise the PO come from VTDManualTest."
    Lamp1 (62,104 30x30), variable: GVL_HMI_VTD.stPdStatus.bCommunicationOk, style: Lamp-Lamp1-Green
    Rectangle (101,104 243x30), "Communication OK"
    Lamp1 (62,138 30x30), variable: GVL_HMI_VTD.stPdStatus.bWcStateError, style: Lamp-Lamp1-Red
    Rectangle (101,138 243x30), "WcState error"
    Rectangle (358,104 146x30), "EtherCAT state"
    Rectangle (504,104 126x30), "%d", text variable: GVL_HMI_VTD.stPdStatus.uiEcState
    Rectangle (358,138 146x30), "PI change counter"
    Rectangle (504,138 126x30), "%u", text variable: GVL_HMI_VTD.stPdStatus.udiInputChangeCount
    Rectangle (63,172 572x28), "EtherCAT state 8 = OP. The counter must keep rising while the drive is powered."
    Rectangle (63,242 58x25), "Word"
    Rectangle (126,242 252x25), "Meaning (MOVISUITE)"
    Rectangle (387,242 117x25), "Raw (hex)"
    Rectangle (514,242 121x25), "Decoded"
    Rectangle (63,272 58x32), "PI 1"
    Rectangle (126,272 252x32), "Status word"
    Rectangle (387,272 117x32), "%04X", text variable: GVL_HMI_VTD.stPdStatus.aProcessInputRaw[1]
    Rectangle (514,272 121x32), "%04X", text variable: GVL_HMI_VTD.stPdStatus.wStatusWord
    Rectangle (63,314 58x32), "PI 2"
    Rectangle (126,314 252x32), "Actual speed"
    Rectangle (387,314 117x32), "%04X", text variable: GVL_HMI_VTD.stPdStatus.aProcessInputRaw[2]
    Rectangle (514,314 121x32), "%d", text variable: GVL_HMI_VTD.stPdStatus.iActualSpeedRaw
    Rectangle (63,356 58x32), "PI 3"
    Rectangle (126,356 252x32), "Status/main fault - subfault"
    Rectangle (387,356 117x32), "%04X", text variable: GVL_HMI_VTD.stPdStatus.aProcessInputRaw[3]
    Rectangle (514,356 121x32), "%04X", text variable: GVL_HMI_VTD.stPdStatus.wFaultCode
    Rectangle (63,398 58x32), "PI 4"
    Rectangle (126,398 252x32), "Torque"
    Rectangle (387,398 117x32), "%04X", text variable: GVL_HMI_VTD.stPdStatus.aProcessInputRaw[4]
    Rectangle (514,398 121x32), "%d", text variable: GVL_HMI_VTD.stPdStatus.iTorqueRaw
    Rectangle (63,440 58x32), "PI 5"
    Rectangle (126,440 252x32), "Digital inputs"
    Rectangle (387,440 117x32), "%04X", text variable: GVL_HMI_VTD.stPdStatus.aProcessInputRaw[5]
    Rectangle (514,440 121x32), "%04X", text variable: GVL_HMI_VTD.stPdStatus.wDigitalInputs
    Rectangle (63,482 58x32), "PI 6"
    Rectangle (126,482 252x32), "Actual application mode"
    Rectangle (387,482 117x32), "%04X", text variable: GVL_HMI_VTD.stPdStatus.aProcessInputRaw[6]
    Rectangle (514,482 121x32), "%u", text variable: GVL_HMI_VTD.stPdStatus.uiActualApplicationMode
    Rectangle (63,524 58x32), "PI 7"
    Rectangle (126,524 252x32), "Actual position - high word"
    Rectangle (387,524 117x32), "%04X", text variable: GVL_HMI_VTD.stPdStatus.aProcessInputRaw[7]
    Rectangle (514,524 121x32), "%d", text variable: GVL_HMI_VTD.stPdStatus.diActualPositionRaw
    Rectangle (63,566 58x32), "PI 8"
    Rectangle (126,566 252x32), "Actual position - low word"
    Rectangle (387,566 117x32), "%04X", text variable: GVL_HMI_VTD.stPdStatus.aProcessInputRaw[8]
    Rectangle (514,566 121x32), "(PI 7 + PI 8)"
    Rectangle (63,610 126x30), "Actual mode"
    Rectangle (193,610 442x30), "%s", text variable: GVL_HMI_VTD.stPdStatus.sActualModeName
    Rectangle (63,650 572x28), "Speed, ramps and position in user units (scaling from MOVISUITE)."
    Rectangle (63,680 572x28), "Torque PI 4 in 0.1 % of nominal motor torque."
    Rectangle (63,710 572x28), "PI 3: high byte = fault, low byte = subfault (active FCB if no fault)."
    Rectangle (688,104 291x56), "%d", text variable: GVL_HMI_VTD.stPdStatus.diActualPositionRaw
    Rectangle (994,104 261x28), "Raw user units"
    Rectangle (994,132 261x28), "Scaling from MOVISUITE"
    Lamp1 (686,206 20x20), variable: GVL_HMI_VTD.stPdStatus.wStatusWord.0, style: Lamp-Lamp1-Green
    Rectangle (713,205 262x22), "0 - Ready"
    Lamp1 (686,229 20x20), variable: GVL_HMI_VTD.stPdStatus.wStatusWord.1, style: Lamp-Lamp1-Green
    Rectangle (713,228 262x22), "1 - STO inactive"
    Lamp1 (686,252 20x20), variable: GVL_HMI_VTD.stPdStatus.wStatusWord.2, style: Lamp-Lamp1-Green
    Rectangle (713,251 262x22), "2 - Output stage enabled"
    Lamp1 (686,275 20x20), variable: GVL_HMI_VTD.stPdStatus.wStatusWord.3, style: Lamp-Lamp1-Green
    Rectangle (713,274 262x22), "3 - Brake released"
    Lamp1 (686,298 20x20), variable: GVL_HMI_VTD.stPdStatus.wStatusWord.4, style: Lamp-Lamp1-Green
    Rectangle (713,297 262x22), "4 - Motor turning"
    Lamp1 (686,321 20x20), variable: GVL_HMI_VTD.stPdStatus.wStatusWord.5, style: Lamp-Lamp1-Green
    Rectangle (713,320 262x22), "5 - Referenced"
    Lamp1 (686,344 20x20), variable: GVL_HMI_VTD.stPdStatus.wStatusWord.6, style: Lamp-Lamp1-Green
    Rectangle (713,343 262x22), "6 - New relative position applied"
    Lamp1 (686,367 20x20), variable: GVL_HMI_VTD.stPdStatus.wStatusWord.7, style: Lamp-Lamp1-Green
    Rectangle (713,366 262x22), "7 - In position"
    Lamp1 (977,206 20x20), variable: GVL_HMI_VTD.stPdStatus.wStatusWord.8, style: Lamp-Lamp1-Red
    Rectangle (1004,205 262x22), "8 - Error"
    Lamp1 (977,229 20x20), variable: GVL_HMI_VTD.stPdStatus.wStatusWord.9, style: Lamp-Lamp1-Yellow
    Rectangle (1004,228 262x22), "9 - Warning"
    Lamp1 (977,252 20x20), variable: GVL_HMI_VTD.stPdStatus.wStatusWord.10, style: Lamp-Lamp1-Green
    Rectangle (1004,251 262x22), "10 - Drive train 2 active"
    Lamp1 (977,275 20x20), variable: GVL_HMI_VTD.stPdStatus.wStatusWord.11, style: Lamp-Lamp1-Green
    Rectangle (1004,274 262x22), "11 - Speed reached"
    Lamp1 (977,298 20x20), variable: GVL_HMI_VTD.stPdStatus.wStatusWord.12, style: Lamp-Lamp1-Green
    Rectangle (1004,297 262x22), "12 - SW limit switches inactive"
    Lamp1 (977,321 20x20), variable: GVL_HMI_VTD.stPdStatus.wStatusWord.13, style: Lamp-Lamp1-Green
    Rectangle (1004,320 262x22), "13 - Reserved"
    Lamp1 (977,344 20x20), variable: GVL_HMI_VTD.stPdStatus.wStatusWord.14, style: Lamp-Lamp1-Green
    Rectangle (1004,343 262x22), "14 - Standby active"
    Lamp1 (977,367 20x20), variable: GVL_HMI_VTD.stPdStatus.wStatusWord.15, style: Lamp-Lamp1-Green
    Rectangle (1004,366 262x22), "15 - Handshake Out"
    Lamp1 (686,424 30x30), variable: GVL_HMI_VTD.stPdStatus.wDigitalInputs.0, style: Lamp-Lamp1-Yellow
    Rectangle (686,456 29x20), "0"
    Lamp1 (722,424 30x30), variable: GVL_HMI_VTD.stPdStatus.wDigitalInputs.1, style: Lamp-Lamp1-Yellow
    Rectangle (722,456 29x20), "1"
    Lamp1 (757,424 30x30), variable: GVL_HMI_VTD.stPdStatus.wDigitalInputs.2, style: Lamp-Lamp1-Yellow
    Rectangle (758,456 29x20), "2"
    Lamp1 (793,424 30x30), variable: GVL_HMI_VTD.stPdStatus.wDigitalInputs.3, style: Lamp-Lamp1-Yellow
    Rectangle (794,456 29x20), "3"
    Lamp1 (829,424 30x30), variable: GVL_HMI_VTD.stPdStatus.wDigitalInputs.4, style: Lamp-Lamp1-Yellow
    Rectangle (830,456 29x20), "4"
    Lamp1 (865,424 30x30), variable: GVL_HMI_VTD.stPdStatus.wDigitalInputs.5, style: Lamp-Lamp1-Yellow
    Rectangle (866,456 29x20), "5"
    Lamp1 (901,424 30x30), variable: GVL_HMI_VTD.stPdStatus.wDigitalInputs.6, style: Lamp-Lamp1-Yellow
    Rectangle (901,456 30x20), "6"
    Lamp1 (937,424 30x30), variable: GVL_HMI_VTD.stPdStatus.wDigitalInputs.7, style: Lamp-Lamp1-Yellow
    Rectangle (937,456 29x20), "7"
    Lamp1 (973,424 30x30), variable: GVL_HMI_VTD.stPdStatus.wDigitalInputs.8, style: Lamp-Lamp1-Yellow
    Rectangle (973,456 29x20), "8"
    Lamp1 (1009,424 30x30), variable: GVL_HMI_VTD.stPdStatus.wDigitalInputs.9, style: Lamp-Lamp1-Yellow
    Rectangle (1009,456 29x20), "9"
    Lamp1 (1045,424 30x30), variable: GVL_HMI_VTD.stPdStatus.wDigitalInputs.10, style: Lamp-Lamp1-Yellow
    Rectangle (1045,456 29x20), "10"
    Lamp1 (1080,424 30x30), variable: GVL_HMI_VTD.stPdStatus.wDigitalInputs.11, style: Lamp-Lamp1-Yellow
    Rectangle (1081,456 29x20), "11"
    Lamp1 (1116,424 30x30), variable: GVL_HMI_VTD.stPdStatus.wDigitalInputs.12, style: Lamp-Lamp1-Yellow
    Rectangle (1117,456 29x20), "12"
    Lamp1 (1152,424 30x30), variable: GVL_HMI_VTD.stPdStatus.wDigitalInputs.13, style: Lamp-Lamp1-Yellow
    Rectangle (1153,456 29x20), "13"
    Lamp1 (1188,424 30x30), variable: GVL_HMI_VTD.stPdStatus.wDigitalInputs.14, style: Lamp-Lamp1-Yellow
    Rectangle (1189,456 29x20), "14"
    Lamp1 (1224,424 30x30), variable: GVL_HMI_VTD.stPdStatus.wDigitalInputs.15, style: Lamp-Lamp1-Yellow
    Rectangle (1224,456 30x20), "15"
    Button (688,514 165x34), "Write enable", colour toggle: GVL_HMI_VTD.stPdCommand.bTestWriteEnable
        toggle GVL_HMI_VTD.stPdCommand.bTestWriteEnable
    Button (863,514 213x34), "Allow control word (PO 1)", colour toggle: GVL_HMI_VTD.stPdCommand.bTestAllowControlWord, input disabled if: NOT GVL_HMI_VTD.stPdCommand.bTestWriteEnable
        toggle GVL_HMI_VTD.stPdCommand.bTestAllowControlWord
    Rectangle (1086,514 169x34), "Elapsed %t[mm:ss]", text variable: GVL_HMI_VTD.stPdStatus.tTestWriteElapsed
    Lamp1 (688,554 30x28), variable: GVL_HMI_VTD.stPdStatus.bTestWriteActive, style: Lamp-Lamp1-Yellow
    Rectangle (722,554 194x28), "Test write active"
    Lamp1 (920,554 30x28), variable: GVL_HMI_VTD.stPdStatus.bTestWriteExpired, style: Lamp-Lamp1-Red
    Rectangle (955,554 300x28), "Timeout expired - toggle Write enable"
    Rectangle (688,590 44x24), "Word"
    Rectangle (735,590 121x24), "Meaning"
    Rectangle (859,590 53x24), "Test"
    Rectangle (915,590 53x24), "Sent"
    Rectangle (688,618 44x32), "PO 1"
    Rectangle (735,618 121x32), "Control word"
    Textfield (859,618 53x32), "%u", text variable: GVL_HMI_VTD.stPdCommand.aTestProcessOutput[1], input disabled if: NOT GVL_HMI_VTD.stPdCommand.bTestAllowControlWord
        OnMouseClick: write the text variable via VisuDialogs.Numpad, min 0, max 65535
    Rectangle (915,618 53x32), "%04X", text variable: GVL_HMI_VTD.stPdStatus.aProcessOutputSent[1]
    Rectangle (688,660 44x32), "PO 2"
    Rectangle (735,660 121x32), "Setpoint speed"
    Textfield (859,660 53x32), "%u", text variable: GVL_HMI_VTD.stPdCommand.aTestProcessOutput[2]
        OnMouseClick: write the text variable via VisuDialogs.Numpad, min 0, max 65535
    Rectangle (915,660 53x32), "%04X", text variable: GVL_HMI_VTD.stPdStatus.aProcessOutputSent[2]
    Rectangle (688,702 44x32), "PO 3"
    Rectangle (735,702 121x32), "Setpoint accel."
    Textfield (859,702 53x32), "%u", text variable: GVL_HMI_VTD.stPdCommand.aTestProcessOutput[3]
        OnMouseClick: write the text variable via VisuDialogs.Numpad, min 0, max 65535
    Rectangle (915,702 53x32), "%04X", text variable: GVL_HMI_VTD.stPdStatus.aProcessOutputSent[3]
    Rectangle (688,744 44x32), "PO 4"
    Rectangle (735,744 121x32), "Setpoint decel."
    Textfield (859,744 53x32), "%u", text variable: GVL_HMI_VTD.stPdCommand.aTestProcessOutput[4]
        OnMouseClick: write the text variable via VisuDialogs.Numpad, min 0, max 65535
    Rectangle (915,744 53x32), "%04X", text variable: GVL_HMI_VTD.stPdStatus.aProcessOutputSent[4]
    Rectangle (974,590 44x24), "Word"
    Rectangle (1021,590 121x24), "Meaning"
    Rectangle (1145,590 53x24), "Test"
    Rectangle (1201,590 53x24), "Sent"
    Rectangle (974,618 44x32), "PO 5"
    Rectangle (1021,618 121x32), "Digital outputs"
    Textfield (1145,618 53x32), "%u", text variable: GVL_HMI_VTD.stPdCommand.aTestProcessOutput[5]
        OnMouseClick: write the text variable via VisuDialogs.Numpad, min 0, max 65535
    Rectangle (1201,618 53x32), "%04X", text variable: GVL_HMI_VTD.stPdStatus.aProcessOutputSent[5]
    Rectangle (974,660 44x32), "PO 6"
    Rectangle (1021,660 121x32), "Setpoint appl. mode"
    Textfield (1145,660 53x32), "%u", text variable: GVL_HMI_VTD.stPdCommand.aTestProcessOutput[6]
        OnMouseClick: write the text variable via VisuDialogs.Numpad, min 0, max 65535
    Rectangle (1201,660 53x32), "%04X", text variable: GVL_HMI_VTD.stPdStatus.aProcessOutputSent[6]
    Rectangle (974,702 44x32), "PO 7"
    Rectangle (1021,702 121x32), "Target pos. high"
    Textfield (1145,702 53x32), "%u", text variable: GVL_HMI_VTD.stPdCommand.aTestProcessOutput[7]
        OnMouseClick: write the text variable via VisuDialogs.Numpad, min 0, max 65535
    Rectangle (1201,702 53x32), "%04X", text variable: GVL_HMI_VTD.stPdStatus.aProcessOutputSent[7]
    Rectangle (974,744 44x32), "PO 8"
    Rectangle (1021,744 121x32), "Target pos. low"
    Textfield (1145,744 53x32), "%u", text variable: GVL_HMI_VTD.stPdCommand.aTestProcessOutput[8]
        OnMouseClick: write the text variable via VisuDialogs.Numpad, min 0, max 65535
    Rectangle (1201,744 53x32), "%04X", text variable: GVL_HMI_VTD.stPdStatus.aProcessOutputSent[8]
    Button (1100,9 160x32), ">> Manual test"
        OnMouseClick: change screen: VTDManualTest
    Rectangle (0,0 156x48)
        OnMouseClick: change screen: Main
    Image (8,4 142x42), image: ImagePool.Logo_Spacemaker
        OnMouseClick: change screen: Main
    Rectangle (0,320 40x160)
        OnMouseClick: OpenDialog Dialog=Dialog, OpenModal=True, PositionX=0, PositionY=0
        OnMouseEnter: OpenDialog Dialog=Dialog, OpenModal=True, PositionX=0, PositionY=0
    Image (0,320 40x160), image: ImagePool.Menu_Tab
        OnMouseClick: OpenDialog Dialog=Dialog, OpenModal=True, PositionX=0, PositionY=0
        OnMouseEnter: OpenDialog Dialog=Dialog, OpenModal=True, PositionX=0, PositionY=0
    Button (63,744 220x36), "SAFETY RESET", colour toggle: GVL_HMI_System.stStatus.bSafetyResetActive
        tap GVL_HMI_System.stCommand.bSafetyReset p3779583253=TRUE
END_VISUALIZATION

// ---- VISUs/VISU_Seeds.TcVIS
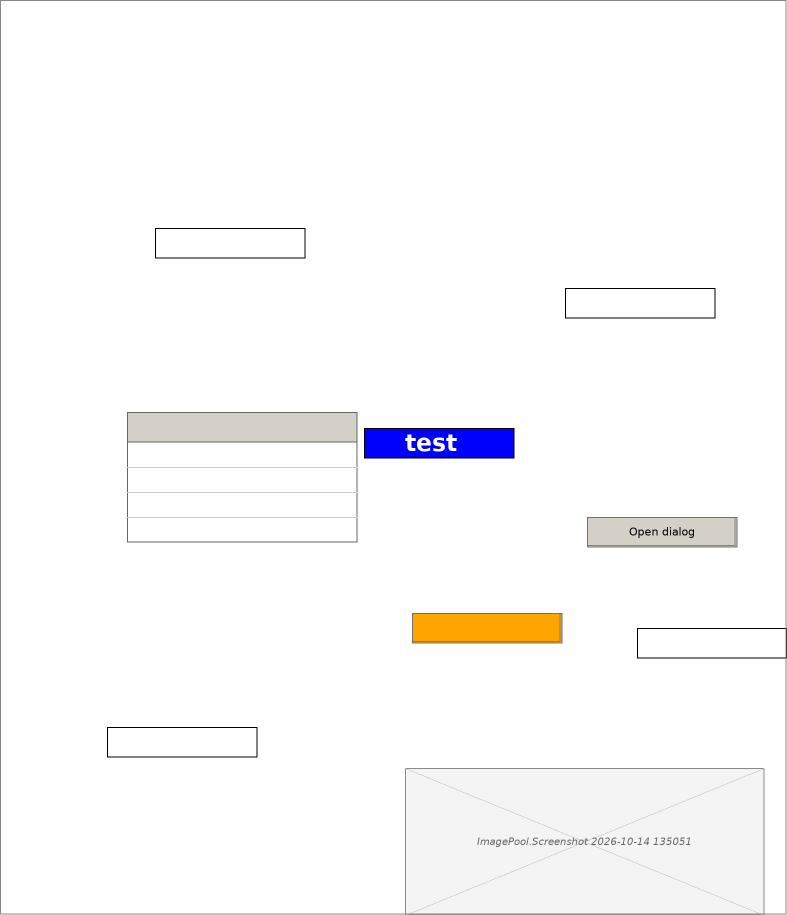
VISUALIZATION VISU_Seeds  // 787x915
    Rectangle (364,428 150x30), "test"
    Button (412,613 150x30)
    Rectangle (565,288 150x30), text list: 'TL_Test'
    Rectangle (637,628 150x30), invisible if: CNV_HMI_IO.HMI_CNV_Backward
    Rectangle (155,228 150x30)
        p2738717112: Control.VTD.Inputs.LE_Position
    Rectangle (107,727 150x30)
        p2277200375: Control.LCnv[1].Inputs.VFD_ActualCurrent
    Image (405,768 359x147), image: ImagePool.Screenshot 2026-10-14 135051
    Frame (453,113 150x30)
        shows FP_Test(bTest := Control.VTD.Docked)
    Table (127,412 230x130), data array: GVL_HMI_VTD.stPdStatus.aProcessInputRaw
        p3854506369: GVL_HMI_VTD.stPdStatus.aProcessInputRaw[INDEX]
        p1014161805: 8 - 1 + INT#1
    Button (587,517 150x30), "Open dialog"
        OnMouseClick: OpenDialog Dialog=Dialog, OpenModal=True, OpenCentered=True
END_VISUALIZATION

// ---- VISUs/VTD.TcVIS
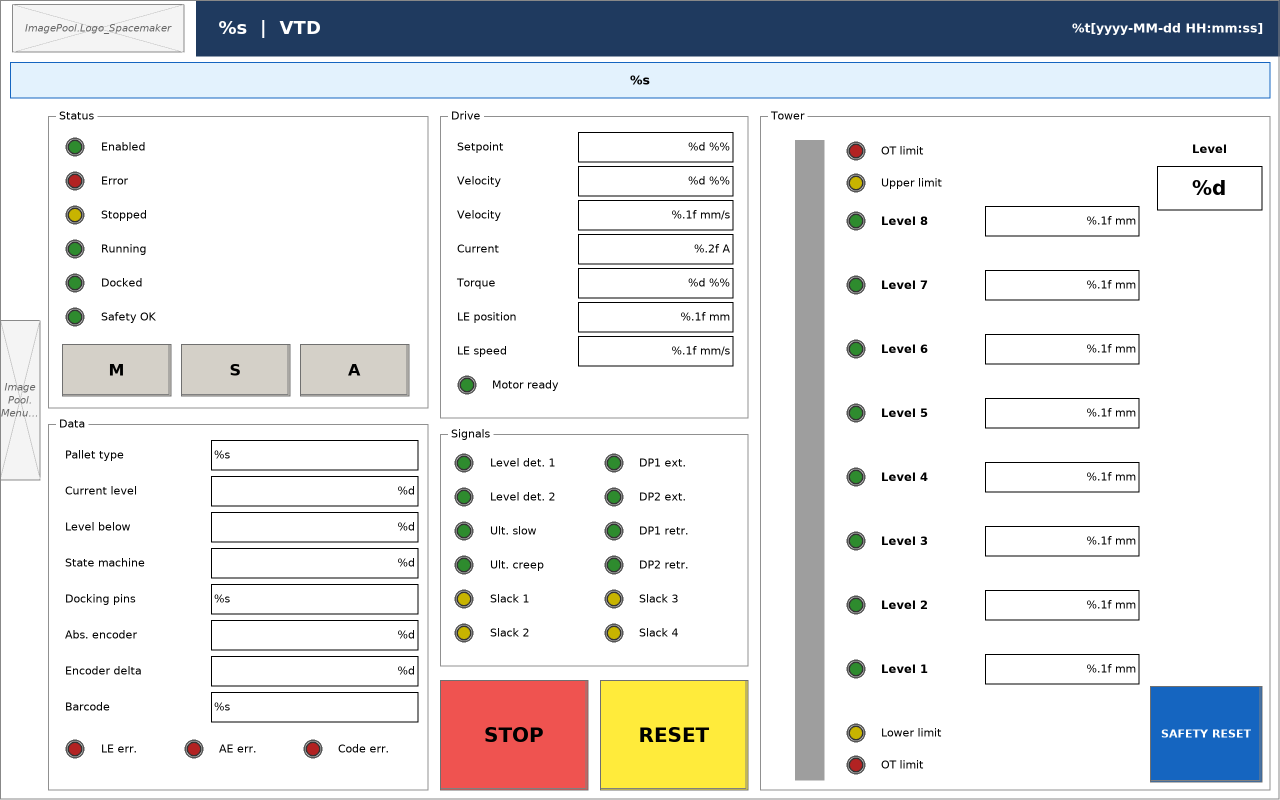
VISUALIZATION VTD  // 1280x800
    Rectangle (0,0 196x56)
        OnMouseClick: change screen: Main
    Image (12,4 172x48), image: ImagePool.Logo_Spacemaker
        OnMouseClick: change screen: Main
    Rectangle (196,0 1084x56), "%s | VTD", text variable: GVL_HMI_System.stStatus.sSystemName
    Rectangle (930,8 336x40), "%t[yyyy-MM-dd HH:mm:ss]", text variable: GVL_HMI_System.stStatus.dtNow
    Rectangle (10,62 1260x36), "%s", text variable: GVL_HMI_System.stStatus.sMessage, colour toggle: GVL_HMI_System.stStatus.bMessageAlarm
    GroupBox (48,108 380x300), "Status"
    Lamp1 (64,136 22x22), variable: GVL_HMI_VTD.stStatus.bEnabled, style: Lamp-Lamp1-Green
    Rectangle (98,132 190x30), "Enabled"
    Lamp1 (64,170 22x22), variable: GVL_HMI_VTD.stStatus.bError, style: Lamp-Lamp1-Red
    Rectangle (98,166 190x30), "Error"
    Lamp1 (64,204 22x22), variable: GVL_HMI_VTD.stStatus.bStopped, style: Lamp-Lamp1-Yellow
    Rectangle (98,200 190x30), "Stopped"
    Lamp1 (64,238 22x22), variable: GVL_HMI_VTD.stStatus.bRunning, style: Lamp-Lamp1-Green
    Rectangle (98,234 190x30), "Running"
    Lamp1 (64,272 22x22), variable: GVL_HMI_VTD.stStatus.bDocked, style: Lamp-Lamp1-Green
    Rectangle (98,268 190x30), "Docked"
    Lamp1 (64,306 22x22), variable: GVL_HMI_VTD.stStatus.bSafetyOk, style: Lamp-Lamp1-Green
    Rectangle (98,302 190x30), "Safety OK"
    Button (62,344 109x52), "M", colour toggle: GVL_HMI_VTD.stStatus.bModeManual
        tap GVL_HMI_VTD.stCommand.bModeManual p3779583253=TRUE
    Button (181,344 109x52), "S", colour toggle: GVL_HMI_VTD.stStatus.bModeSemi
        tap GVL_HMI_VTD.stCommand.bModeSemi p3779583253=TRUE
    Button (300,344 109x52), "A", colour toggle: GVL_HMI_VTD.stStatus.bModeAuto
        tap GVL_HMI_VTD.stCommand.bModeAuto p3779583253=TRUE
    GroupBox (48,416 380x374), "Data"
    Rectangle (62,440 143x30), "Pallet type"
    Rectangle (211,440 207x30), "%s", text variable: GVL_HMI_VTD.stStatus.sPalletType
    Rectangle (62,476 143x30), "Current level"
    Rectangle (211,476 207x30), "%d", text variable: GVL_HMI_VTD.stStatus.uiCurrentLevel
    Rectangle (62,512 143x30), "Level below"
    Rectangle (211,512 207x30), "%d", text variable: GVL_HMI_VTD.stStatus.uiLevelBelow
    Rectangle (62,548 143x30), "State machine"
    Rectangle (211,548 207x30), "%d", text variable: GVL_HMI_VTD.stStatus.uiStateMachine
    Rectangle (62,584 143x30), "Docking pins"
    Rectangle (211,584 207x30), "%s", text variable: GVL_HMI_VTD.stStatus.sDockingPinState
    Rectangle (62,620 143x30), "Abs. encoder"
    Rectangle (211,620 207x30), "%d", text variable: GVL_HMI_VTD.stStatus.diAbsoluteEncoder
    Rectangle (62,656 143x30), "Encoder delta"
    Rectangle (211,656 207x30), "%d", text variable: GVL_HMI_VTD.stStatus.iEncoderDelta
    Rectangle (62,692 143x30), "Barcode"
    Rectangle (211,692 207x30), "%s", text variable: GVL_HMI_VTD.stStatus.sBarcode
    Lamp1 (64,738 22x22), variable: GVL_HMI_VTD.stStatus.bLinearEncoderError, style: Lamp-Lamp1-Red
    Rectangle (98,734 78x30), "LE err."
    Lamp1 (183,738 22x22), variable: GVL_HMI_VTD.stStatus.bAbsoluteEncoderError, style: Lamp-Lamp1-Red
    Rectangle (216,734 79x30), "AE err."
    Lamp1 (302,738 22x22), variable: GVL_HMI_VTD.stStatus.bBarcodeError, style: Lamp-Lamp1-Red
    Rectangle (335,734 78x30), "Code err."
    GroupBox (440,108 308x310), "Drive"
    Rectangle (454,132 118x30), "Setpoint"
    Rectangle (578,132 155x30), "%d %%", text variable: GVL_HMI_VTD.stStatus.iSetpoint_pct
    Rectangle (454,166 118x30), "Velocity"
    Rectangle (578,166 155x30), "%d %%", text variable: GVL_HMI_VTD.stStatus.iVelocity_pct
    Rectangle (454,200 118x30), "Velocity"
    Rectangle (578,200 155x30), "%.1f mm/s", text variable: GVL_HMI_VTD.stStatus.rVelocity_mm_s
    Rectangle (454,234 118x30), "Current"
    Rectangle (578,234 155x30), "%.2f A", text variable: GVL_HMI_VTD.stStatus.rCurrent_A
    Rectangle (454,268 118x30), "Torque"
    Rectangle (578,268 155x30), "%d %%", text variable: GVL_HMI_VTD.stStatus.iTorque_pct
    Rectangle (454,302 118x30), "LE position"
    Rectangle (578,302 155x30), "%.1f mm", text variable: GVL_HMI_VTD.stStatus.rLePosition_mm
    Rectangle (454,336 118x30), "LE speed"
    Rectangle (578,336 155x30), "%.1f mm/s", text variable: GVL_HMI_VTD.stStatus.rLeSpeed_mm_s
    Lamp1 (456,374 22x22), variable: GVL_HMI_VTD.stStatus.bMotorReady, style: Lamp-Lamp1-Green
    Rectangle (489,370 190x30), "Motor ready"
    GroupBox (440,426 308x240), "Signals"
    Lamp1 (453,452 22x22), variable: GVL_HMI_VTD.stStatus.bLevelDetect1, style: Lamp-Lamp1-Green
    Rectangle (487,448 109x30), "Level det. 1"
    Lamp1 (453,486 22x22), variable: GVL_HMI_VTD.stStatus.bLevelDetect2, style: Lamp-Lamp1-Green
    Rectangle (487,482 109x30), "Level det. 2"
    Lamp1 (453,520 22x22), variable: GVL_HMI_VTD.stStatus.bUltimateSlowdown, style: Lamp-Lamp1-Green
    Rectangle (487,516 109x30), "Ult. slow"
    Lamp1 (453,554 22x22), variable: GVL_HMI_VTD.stStatus.bUltimateCreep, style: Lamp-Lamp1-Green
    Rectangle (487,550 109x30), "Ult. creep"
    Lamp1 (453,588 22x22), variable: GVL_HMI_VTD.stStatus.abChainSlack[1], style: Lamp-Lamp1-Yellow
    Rectangle (487,584 109x30), "Slack 1"
    Lamp1 (453,622 22x22), variable: GVL_HMI_VTD.stStatus.abChainSlack[2], style: Lamp-Lamp1-Yellow
    Rectangle (487,618 109x30), "Slack 2"
    Lamp1 (603,452 22x22), variable: GVL_HMI_VTD.stStatus.bDp1Extended, style: Lamp-Lamp1-Green
    Rectangle (636,448 110x30), "DP1 ext."
    Lamp1 (603,486 22x22), variable: GVL_HMI_VTD.stStatus.bDp2Extended, style: Lamp-Lamp1-Green
    Rectangle (636,482 110x30), "DP2 ext."
    Lamp1 (603,520 22x22), variable: GVL_HMI_VTD.stStatus.bDp1Retracted, style: Lamp-Lamp1-Green
    Rectangle (636,516 110x30), "DP1 retr."
    Lamp1 (603,554 22x22), variable: GVL_HMI_VTD.stStatus.bDp2Retracted, style: Lamp-Lamp1-Green
    Rectangle (636,550 110x30), "DP2 retr."
    Lamp1 (603,588 22x22), variable: GVL_HMI_VTD.stStatus.abChainSlack[3], style: Lamp-Lamp1-Yellow
    Rectangle (636,584 110x30), "Slack 3"
    Lamp1 (603,622 22x22), variable: GVL_HMI_VTD.stStatus.abChainSlack[4], style: Lamp-Lamp1-Yellow
    Rectangle (636,618 110x30), "Slack 4"
    Button (440,680 148x110), "STOP"
        tap GVL_HMI_VTD.stCommand.bStop p3779583253=TRUE
    Button (600,680 148x110), "RESET"
        tap GVL_HMI_VTD.stCommand.bReset p3779583253=TRUE
    GroupBox (760,108 510x682), "Tower"
    Rectangle (795,140 29x640)
    Lamp1 (845,140 22x22), variable: GVL_HMI_VTD.stStatus.bUpperOvertravel, style: Lamp-Lamp1-Red
    Rectangle (878,136 131x30), "OT limit"
    Lamp1 (845,172 22x22), variable: GVL_HMI_VTD.stStatus.bUpperLimit, style: Lamp-Lamp1-Yellow
    Rectangle (878,168 131x30), "Upper limit"
    Lamp1 (845,210 22x22), variable: GVL_HMI_VTD.stStatus.abLevelReached[8], style: Lamp-Lamp1-Green
    Rectangle (878,206 95x30), "Level 8"
    Rectangle (985,206 154x30), "%.1f mm", text variable: GVL_HMI_VTD.stStatus.arLevelPosition_mm[8]
    Lamp1 (845,274 22x22), variable: GVL_HMI_VTD.stStatus.abLevelReached[7], style: Lamp-Lamp1-Green
    Rectangle (878,270 95x30), "Level 7"
    Rectangle (985,270 154x30), "%.1f mm", text variable: GVL_HMI_VTD.stStatus.arLevelPosition_mm[7]
    Lamp1 (845,338 22x22), variable: GVL_HMI_VTD.stStatus.abLevelReached[6], style: Lamp-Lamp1-Green
    Rectangle (878,334 95x30), "Level 6"
    Rectangle (985,334 154x30), "%.1f mm", text variable: GVL_HMI_VTD.stStatus.arLevelPosition_mm[6]
    Lamp1 (845,402 22x22), variable: GVL_HMI_VTD.stStatus.abLevelReached[5], style: Lamp-Lamp1-Green
    Rectangle (878,398 95x30), "Level 5"
    Rectangle (985,398 154x30), "%.1f mm", text variable: GVL_HMI_VTD.stStatus.arLevelPosition_mm[5]
    Lamp1 (845,466 22x22), variable: GVL_HMI_VTD.stStatus.abLevelReached[4], style: Lamp-Lamp1-Green
    Rectangle (878,462 95x30), "Level 4"
    Rectangle (985,462 154x30), "%.1f mm", text variable: GVL_HMI_VTD.stStatus.arLevelPosition_mm[4]
    Lamp1 (845,530 22x22), variable: GVL_HMI_VTD.stStatus.abLevelReached[3], style: Lamp-Lamp1-Green
    Rectangle (878,526 95x30), "Level 3"
    Rectangle (985,526 154x30), "%.1f mm", text variable: GVL_HMI_VTD.stStatus.arLevelPosition_mm[3]
    Lamp1 (845,594 22x22), variable: GVL_HMI_VTD.stStatus.abLevelReached[2], style: Lamp-Lamp1-Green
    Rectangle (878,590 95x30), "Level 2"
    Rectangle (985,590 154x30), "%.1f mm", text variable: GVL_HMI_VTD.stStatus.arLevelPosition_mm[2]
    Lamp1 (845,658 22x22), variable: GVL_HMI_VTD.stStatus.abLevelReached[1], style: Lamp-Lamp1-Green
    Rectangle (878,654 95x30), "Level 1"
    Rectangle (985,654 154x30), "%.1f mm", text variable: GVL_HMI_VTD.stStatus.arLevelPosition_mm[1]
    Lamp1 (845,722 22x22), variable: GVL_HMI_VTD.stStatus.bLowerLimit, style: Lamp-Lamp1-Yellow
    Rectangle (878,718 131x30), "Lower limit"
    Lamp1 (845,754 22x22), variable: GVL_HMI_VTD.stStatus.bLowerOvertravel, style: Lamp-Lamp1-Red
    Rectangle (878,750 131x30), "OT limit"
    Rectangle (1157,136 105x26), "Level"
    Rectangle (1157,166 105x44), "%d", text variable: GVL_HMI_VTD.stStatus.uiCurrentLevel
    Rectangle (0,320 40x160)
        OnMouseClick: OpenDialog Dialog=Dialog, OpenModal=True, PositionX=0, PositionY=0
        OnMouseEnter: OpenDialog Dialog=Dialog, OpenModal=True, PositionX=0, PositionY=0
    Image (0,320 40x160), image: ImagePool.Menu_Tab
        OnMouseClick: OpenDialog Dialog=Dialog, OpenModal=True, PositionX=0, PositionY=0
        OnMouseEnter: OpenDialog Dialog=Dialog, OpenModal=True, PositionX=0, PositionY=0
    Button (1150,686 112x96), "SAFETY RESET", colour toggle: GVL_HMI_System.stStatus.bSafetyResetActive
        tap GVL_HMI_System.stCommand.bSafetyReset p3779583253=TRUE
END_VISUALIZATION

// ---- VISUs/VTDManualTest.TcVIS
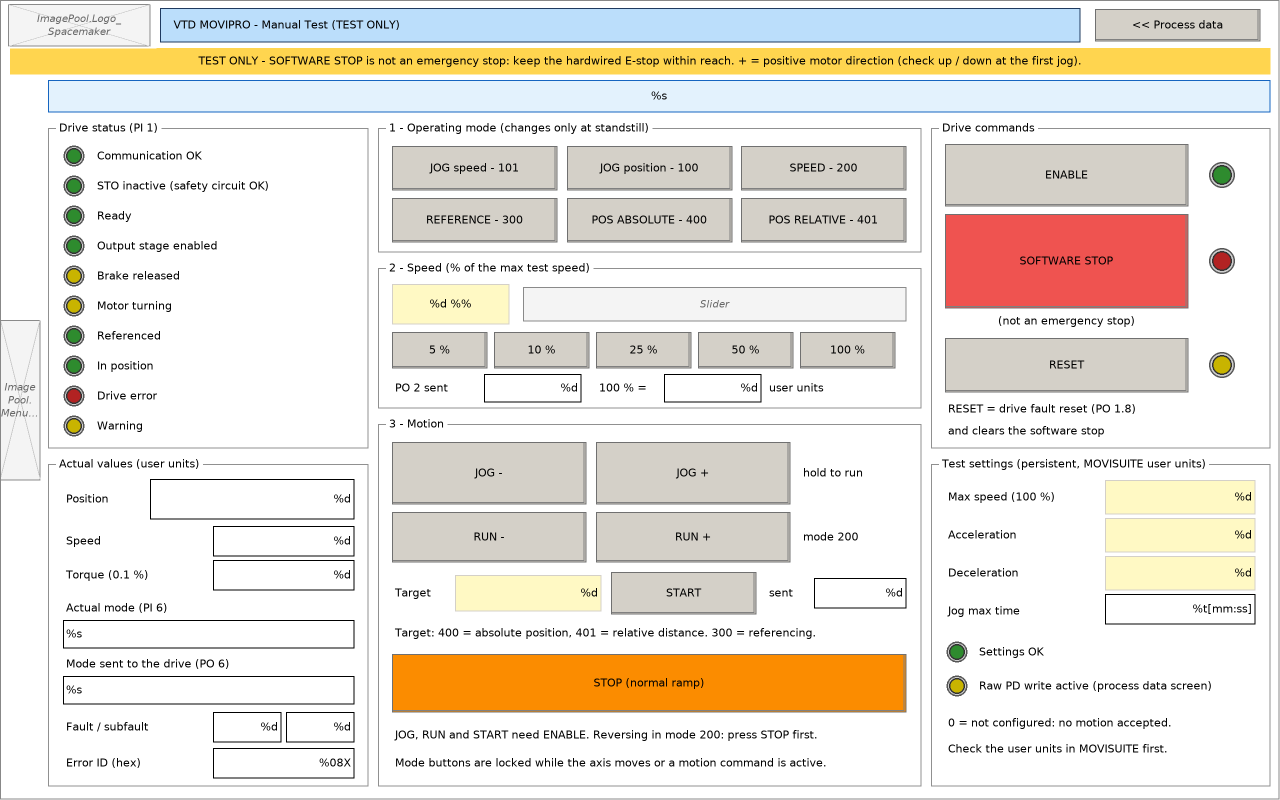
VISUALIZATION VTDManualTest  // 1280x800
    Rectangle (160,8 920x34), "VTD MOVIPRO - Manual Test (TEST ONLY)"
    Button (1095,9 165x32), "<< Process data"
        OnMouseClick: change screen: Visualization
    Rectangle (10,48 1260x26), "TEST ONLY - SOFTWARE STOP is not an emergency stop: keep the hardwired E-stop within reach. + = positive motor direction (check up / down at the first jog)."
    Rectangle (48,80 1222x32), "%s", text variable: GVL_HMI_VTD.stManualStatus.sMessage, colour toggle: GVL_HMI_VTD.stManualStatus.bMessageAlarm
    GroupBox (48,120 320x328), "Drive status (PI 1)"
    Lamp1 (62,144 24x24), variable: GVL_HMI_VTD.stManualStatus.stDrive.bCommunicationOk, style: Lamp-Lamp1-Green
    Rectangle (94,142 261x28), "Communication OK"
    Lamp1 (62,174 24x24), variable: GVL_HMI_VTD.stManualStatus.stDrive.bStoInactive, style: Lamp-Lamp1-Green
    Rectangle (94,172 261x28), "STO inactive (safety circuit OK)"
    Lamp1 (62,204 24x24), variable: GVL_HMI_VTD.stManualStatus.stDrive.bReady, style: Lamp-Lamp1-Green
    Rectangle (94,202 261x28), "Ready"
    Lamp1 (62,234 24x24), variable: GVL_HMI_VTD.stManualStatus.stDrive.bOutputStageEnabled, style: Lamp-Lamp1-Green
    Rectangle (94,232 261x28), "Output stage enabled"
    Lamp1 (62,264 24x24), variable: GVL_HMI_VTD.stManualStatus.stDrive.bBrakeReleased, style: Lamp-Lamp1-Yellow
    Rectangle (94,262 261x28), "Brake released"
    Lamp1 (62,294 24x24), variable: GVL_HMI_VTD.stManualStatus.stDrive.bMotorTurning, style: Lamp-Lamp1-Yellow
    Rectangle (94,292 261x28), "Motor turning"
    Lamp1 (62,324 24x24), variable: GVL_HMI_VTD.stManualStatus.stDrive.bReferenced, style: Lamp-Lamp1-Green
    Rectangle (94,322 261x28), "Referenced"
    Lamp1 (62,354 24x24), variable: GVL_HMI_VTD.stManualStatus.stDrive.bInPosition, style: Lamp-Lamp1-Green
    Rectangle (94,352 261x28), "In position"
    Lamp1 (62,384 24x24), variable: GVL_HMI_VTD.stManualStatus.stDrive.bError, style: Lamp-Lamp1-Red
    Rectangle (94,382 261x28), "Drive error"
    Lamp1 (62,414 24x24), variable: GVL_HMI_VTD.stManualStatus.stDrive.bWarning, style: Lamp-Lamp1-Yellow
    Rectangle (94,412 261x28), "Warning"
    GroupBox (48,456 320x330), "Actual values (user units)"
    Rectangle (63,484 82x30), "Position"
    Rectangle (150,479 204x40), "%d", text variable: GVL_HMI_VTD.stManualStatus.stDrive.diActualPosition
    Rectangle (63,526 145x30), "Speed"
    Rectangle (213,526 141x30), "%d", text variable: GVL_HMI_VTD.stManualStatus.stDrive.iActualSpeed
    Rectangle (63,560 145x30), "Torque (0.1 %)"
    Rectangle (213,560 141x30), "%d", text variable: GVL_HMI_VTD.stManualStatus.stDrive.iActualTorque_0p1pct
    Rectangle (63,596 291x24), "Actual mode (PI 6)"
    Rectangle (63,620 291x28), "%s", text variable: GVL_HMI_VTD.stManualStatus.sActualModeName
    Rectangle (63,652 291x24), "Mode sent to the drive (PO 6)"
    Rectangle (63,676 291x28), "%s", text variable: GVL_HMI_VTD.stManualStatus.sModeActiveName
    Rectangle (63,712 145x30), "Fault / subfault"
    Rectangle (213,712 68x30), "%d", text variable: GVL_HMI_VTD.stManualStatus.stDrive.byFaultCode
    Rectangle (286,712 68x30), "%d", text variable: GVL_HMI_VTD.stManualStatus.stDrive.bySubfaultCode
    Rectangle (63,748 145x30), "Error ID (hex)"
    Rectangle (213,748 141x30), "%08X", text variable: GVL_HMI_VTD.stManualStatus.udiErrorId
    GroupBox (378,120 543x132), "1 - Operating mode (changes only at standstill)"
    Button (392,146 165x44), "JOG speed - 101", colour toggle: GVL_HMI_VTD.stManualStatus.bModeJogSpeed, input disabled if: NOT GVL_HMI_VTD.stManualStatus.bModeChangeAllowed
        OnMouseClick: execute { GVL_HMI_VTD.stManualCommand.eModeRequest := E_SEW_MovikitMode.JogSpeedControlled; }
    Button (567,146 165x44), "JOG position - 100", colour toggle: GVL_HMI_VTD.stManualStatus.bModeJogPosition, input disabled if: NOT GVL_HMI_VTD.stManualStatus.bModeChangeAllowed
        OnMouseClick: execute { GVL_HMI_VTD.stManualCommand.eModeRequest := E_SEW_MovikitMode.JogPositionControlled; }
    Button (741,146 165x44), "SPEED - 200", colour toggle: GVL_HMI_VTD.stManualStatus.bModeSpeed, input disabled if: NOT GVL_HMI_VTD.stManualStatus.bModeChangeAllowed
        OnMouseClick: execute { GVL_HMI_VTD.stManualCommand.eModeRequest := E_SEW_MovikitMode.Speed; }
    Button (392,198 165x44), "REFERENCE - 300", colour toggle: GVL_HMI_VTD.stManualStatus.bModeReferencing, input disabled if: NOT GVL_HMI_VTD.stManualStatus.bModeChangeAllowed
        OnMouseClick: execute { GVL_HMI_VTD.stManualCommand.eModeRequest := E_SEW_MovikitMode.ReferencingOffsetConfigured; }
    Button (567,198 165x44), "POS ABSOLUTE - 400", colour toggle: GVL_HMI_VTD.stManualStatus.bModePositionAbsolute, input disabled if: NOT GVL_HMI_VTD.stManualStatus.bModeChangeAllowed
        OnMouseClick: execute { GVL_HMI_VTD.stManualCommand.eModeRequest := E_SEW_MovikitMode.PositioningAbsolute; }
    Button (741,198 165x44), "POS RELATIVE - 401", colour toggle: GVL_HMI_VTD.stManualStatus.bModePositionRelative, input disabled if: NOT GVL_HMI_VTD.stManualStatus.bModeChangeAllowed
        OnMouseClick: execute { GVL_HMI_VTD.stManualCommand.eModeRequest := E_SEW_MovikitMode.PositioningRelative; }
    GroupBox (378,260 543x148), "2 - Speed (% of the max test speed)"
    Textfield (392,284 117x40), "%d %%", text variable: GVL_HMI_VTD.stManualCommand.iSpeedPercent
        OnMouseClick: write the text variable via VisuDialogs.Numpad, min 0, max 100
    Slider (523,287 383x34), variable: GVL_HMI_VTD.stManualCommand.iSpeedPercent, scale 0..100
    Button (392,332 95x36), "5 %"
        OnMouseClick: execute { GVL_HMI_VTD.stManualCommand.iSpeedPercent := 5; }
    Button (494,332 95x36), "10 %"
        OnMouseClick: execute { GVL_HMI_VTD.stManualCommand.iSpeedPercent := 10; }
    Button (596,332 95x36), "25 %"
        OnMouseClick: execute { GVL_HMI_VTD.stManualCommand.iSpeedPercent := 25; }
    Button (698,332 95x36), "50 %"
        OnMouseClick: execute { GVL_HMI_VTD.stManualCommand.iSpeedPercent := 50; }
    Button (800,332 95x36), "100 %"
        OnMouseClick: execute { GVL_HMI_VTD.stManualCommand.iSpeedPercent := 100; }
    Rectangle (392,374 92x28), "PO 2 sent"
    Rectangle (484,374 97x28), "%d", text variable: GVL_HMI_VTD.stManualStatus.iSpeedSetpoint
    Rectangle (596,374 68x28), "100 % ="
    Rectangle (664,374 97x28), "%d", text variable: GVL_HMI_VTD.stManualSettings.iMaxSpeed
    Rectangle (766,374 140x28), "user units"
    GroupBox (378,416 543x370), "3 - Motion"
    Button (392,442 194x62), "JOG -", colour toggle: GVL_HMI_VTD.stManualStatus.bJogNegativeActive, input disabled if: NOT GVL_HMI_VTD.stManualStatus.bJogAvailable
        tap GVL_HMI_VTD.stManualCommand.bJogNegative p3779583253=TRUE
    Button (596,442 194x62), "JOG +", colour toggle: GVL_HMI_VTD.stManualStatus.bJogPositiveActive, input disabled if: NOT GVL_HMI_VTD.stManualStatus.bJogAvailable
        tap GVL_HMI_VTD.stManualCommand.bJogPositive p3779583253=TRUE
    Rectangle (800,458 111x30), "hold to run"
    Button (392,512 194x50), "RUN -", colour toggle: GVL_HMI_VTD.stManualStatus.bRunNegativeActive, input disabled if: NOT GVL_HMI_VTD.stManualStatus.bRunAvailable
        tap GVL_HMI_VTD.stManualCommand.bRunNegative p3779583253=TRUE
    Button (596,512 194x50), "RUN +", colour toggle: GVL_HMI_VTD.stManualStatus.bRunPositiveActive, input disabled if: NOT GVL_HMI_VTD.stManualStatus.bRunAvailable
        tap GVL_HMI_VTD.stManualCommand.bRunPositive p3779583253=TRUE
    Rectangle (800,522 111x30), "mode 200"
    Rectangle (392,578 63x30), "Target"
    Textfield (455,575 146x36), "%d", text variable: GVL_HMI_VTD.stManualCommand.diTargetPosition
        OnMouseClick: write the text variable via VisuDialogs.Numpad, min -2147483648, max 2147483647
    Button (611,572 145x42), "START", colour toggle: GVL_HMI_VTD.stManualStatus.bStartActive, input disabled if: NOT GVL_HMI_VTD.stManualStatus.bStartAvailable
        tap GVL_HMI_VTD.stManualCommand.bStart p3779583253=TRUE
    Rectangle (766,578 48x30), "sent"
    Rectangle (814,578 92x30), "%d", text variable: GVL_HMI_VTD.stManualStatus.diTargetPositionSent
    Rectangle (392,620 514x26), "Target: 400 = absolute position, 401 = relative distance. 300 = referencing."
    Button (392,654 514x58), "STOP (normal ramp)"
        tap GVL_HMI_VTD.stManualCommand.bStop p3779583253=TRUE
    Rectangle (392,722 514x26), "JOG, RUN and START need ENABLE. Reversing in mode 200: press STOP first."
    Rectangle (392,750 514x26), "Mode buttons are locked while the axis moves or a motion command is active."
    GroupBox (931,120 339x328), "Drive commands"
    Button (945,144 243x62), "ENABLE", colour toggle: GVL_HMI_VTD.stManualStatus.bEnableActive
        toggle GVL_HMI_VTD.stManualCommand.bEnable
    Lamp1 (1207,160 30x30), variable: GVL_HMI_VTD.stManualStatus.bEnableActive, style: Lamp-Lamp1-Green
    Button (945,214 243x94), "SOFTWARE STOP"
        tap GVL_HMI_VTD.stManualCommand.bSoftwareStop p3779583253=TRUE
    Lamp1 (1207,246 30x30), variable: GVL_HMI_VTD.stManualStatus.bSoftwareStopActive, style: Lamp-Lamp1-Red
    Rectangle (945,310 243x22), "(not an emergency stop)"
    Button (945,338 243x54), "RESET"
        tap GVL_HMI_VTD.stManualCommand.bReset p3779583253=TRUE
    Lamp1 (1207,350 30x30), variable: GVL_HMI_VTD.stManualStatus.bFaultResetActive, style: Lamp-Lamp1-Yellow
    Rectangle (945,398 315x22), "RESET = drive fault reset (PO 1.8)"
    Rectangle (945,420 315x22), "and clears the software stop"
    GroupBox (931,456 339x330), "Test settings (persistent, MOVISUITE user units)"
    Rectangle (945,482 155x30), "Max speed (100 %)"
    Textfield (1105,480 150x34), "%d", text variable: GVL_HMI_VTD.stManualSettings.iMaxSpeed
        OnMouseClick: write the text variable via VisuDialogs.Numpad, min 0, max 32767
    Rectangle (945,520 155x30), "Acceleration"
    Textfield (1105,518 150x34), "%d", text variable: GVL_HMI_VTD.stManualSettings.uiAcceleration
        OnMouseClick: write the text variable via VisuDialogs.Numpad, min 0, max 65535
    Rectangle (945,558 155x30), "Deceleration"
    Textfield (1105,556 150x34), "%d", text variable: GVL_HMI_VTD.stManualSettings.uiDeceleration
        OnMouseClick: write the text variable via VisuDialogs.Numpad, min 0, max 65535
    Rectangle (945,596 155x30), "Jog max time"
    Rectangle (1105,594 150x30), "%t[mm:ss]", text variable: GVL_HMI_VTD.stManualSettings.tJogMaxTime
    Lamp1 (945,640 24x24), variable: GVL_HMI_VTD.stManualStatus.bSettingsValid, style: Lamp-Lamp1-Green
    Rectangle (976,637 281x30), "Settings OK"
    Lamp1 (945,674 24x24), variable: GVL_HMI_VTD.stManualStatus.bRawWriteActive, style: Lamp-Lamp1-Yellow
    Rectangle (976,671 281x30), "Raw PD write active (process data screen)"
    Rectangle (945,710 315x26), "0 = not configured: no motion accepted."
    Rectangle (945,736 315x26), "Check the user units in MOVISUITE first."
    Rectangle (0,0 156x48)
        OnMouseClick: change screen: Main
    Image (8,4 142x42), image: ImagePool.Logo_Spacemaker
        OnMouseClick: change screen: Main
    Rectangle (0,320 40x160)
        OnMouseClick: OpenDialog Dialog=Dialog, OpenModal=True, PositionX=0, PositionY=0
        OnMouseEnter: OpenDialog Dialog=Dialog, OpenModal=True, PositionX=0, PositionY=0
    Image (0,320 40x160), image: ImagePool.Menu_Tab
        OnMouseClick: OpenDialog Dialog=Dialog, OpenModal=True, PositionX=0, PositionY=0
        OnMouseEnter: OpenDialog Dialog=Dialog, OpenModal=True, PositionX=0, PositionY=0
END_VISUALIZATION

// ---- VISUs/VTD_Settings.TcVIS
VISUALIZATION VTD_Settings  // 1024x768
END_VISUALIZATION
